(* IEC 61131-3 sources: daoli-st-library/DL_Process (part 8) *)

(* ---- FB_DL_TruckScaleSeq.st ---- *)
(*==============================================================================
 * 组件名称 (Component)  : FB_DL_TruckScaleSeq
 * 所属子库 (Sublibrary) : DL_Process
 * 当前版本 (Version)    : 1.0.2
 * 兼容性   (Platform)   : CODESYS 3.5 / TwinCAT 3 / 汇川 InoProShop / Machine Expert
 *                         仅依赖 Standard.library + DL_ 库内既有件，零厂商方言
 * 来源标签 (Source)     : self-std
 * 功能描述 (Function)   : 车辆过磅称重流程七态顺控：空载等待 -> 车辆上磅（到位
 *                         开关）-> 稳定窗（称重稳定判据，委托 FB_DL_SignalStatistics
 *                         统计内核，峰峰值 < 容差判稳）-> 读数锁存（皮重 / 毛重
 *                         配对）-> 下磅 -> 台账推进（8 条定长环形，写指针饱和）。
 *                         超时未稳定置码重测；防作弊窗（读数期间磅台扰动检测）；
 *                         毛重 < 皮重（亏吨）显式码不静默取负净重。
 * 委托清单 (Delegation) : FB_DL_SignalStatistics（DL_MathData，稳态窗口径次源，
 *                         实例化组合调用——峰峰值 fRange 即稳定判据核）
 * 配比约束 (R100)       : tStableTimeout 必须大于统计窗填满耗时（nStableSamples ×
 *                         任务周期），否则未满窗即被超时重测，稳定判据永不达成。
 * 遗留假设三句声明 (R95): ①代理值：稳定窗以「样本数 nStableSamples × 任务周期」
 *                         代理时间窗 tStableWin；②覆盖范围：任务周期已知且恒定的
 *                         调用场合；③覆盖不到的区间：任务周期漂移 / 变长场合由
 *                         tStableTimeout 超时重测兜底，最坏表现是判稳变慢而非误判。
 * 边界与语义披露 (Boundary disclosure) :
 *   1) 读数未锁存前下磅（bOnScale 在稳定 / 锁存相消失）-> 流程作废 + 台账不写入
 *      （信息级），统计窗清零重来。
 *   2) 防作弊窗：稳定相内磅台到位信号闪断视为扰动（车未完全上磅 / 人为干预），
 *      置信息级并回稳定相重测，杜绝在扰动读数上锁存。
 *   3) 毛重 < 皮重（亏吨）为显式信息级：净重置 0 出台账，绝不静默取负
 *      （负净重会污染库存对账，R81 还原方向不饱和口径同理）。
 *   4) 皮 / 毛配对以「皮重槽与毛重槽均已锁存」为准，不做车号强校验（车号仅入
 *      台账留痕）；配对完成后双槽清零迎接下一车。
 *   5) 称重值非有限属**运行时信号失效**，不是组态错误：自 v1.0.2 起拆为独立信号闸——
 *      本拍只判 NaN / Inf 并置信息级 16#0005_04DD，统计与判据一律使用上一次有效值
 *      快照（fWeightHold），不锁存、不置 bError、不迁 eFault；失效持续由稳定超时
 *      重测（04D9）兜底。判定拍与消费拍强制错开一拍（本拍判定 -> 下拍消费
 *      bWeightBad），杜绝同拍把脏值锁进皮毛槽。
 *   6) 组态闸（bCfgBad）自 v1.0.2 起只含**静态组态量**（容差 / 超时窗 / 窗样本数），
 *      运行时信号不得进入组态锁存路径（避免一拍 NaN 让磅房永久锁死，R152）。
 * 故障码表 (Error codes) :
 *   16#0005_03B2 [故障级] 稳定窗组态非法（容差 <= 0 / 超时 <= 0 / 窗样本数越域）
 *                 反证：回退后流程照常，码位是组态错误唯一可见出口。
 *   16#0005_04D6 [信息级] 未锁存先下磅，流程作废台账不写入
 *                 反证：作废后回空闲与「正常完成」输出组合不同但作废原因（司机
 *                 误操作 / 磅台故障）不可区分，码位承载事件事实。
 *   16#0005_04D7 [信息级] 亏吨（毛重 < 皮重），净重置 0 出台账
 *                 反证：净重 0 与「空车皮重恰好等于毛重」组合相同，码位区分
 *                 正常零载与亏吨异常。
 *   16#0005_04D8 [信息级] 读数期磅台扰动（防作弊窗触发），重测
 *                 反证：重测与「正常重来」输出组合相同，码位是防作弊事实唯一出口。
 *   16#0005_04D9 [信息级] 超时未稳定，清窗重测
 *                 反证：重测与防作弊重测输出组合相似（均回稳定相），码位区分
 *                 「称量不稳」与「磅台扰动」两种成因（R190）。
 *   16#0005_04DD [信息级] 称重信号非有限（NaN / Inf），保持上次有效值不锁存
 *                 反证：保持时 fWeightHold 不变，与「称重值恰好稳定不变」的输出组合
 *                 完全相同；无码则信号断线被误读为「读数极稳」而照常判稳锁存，
 *                 该误判在现有输出上不可观测（R90 反证成立，R69 点修④）。
 * 码位总账 (Code ledger) : 16#0005_03B2 用 ｜ 16#0005_04D6 / 04D7 / 04D8 / 04D9 / 04DD 用
 * 依赖     (Depends)    : FB_DL_SignalStatistics
 * 红线自检 (Redline)    : R1 ✓ 零全局变量与 VAR_EXTERNAL ｜ R2 ✓ 零 %I/%Q 物理地址
 *                         R3 ✓ 纯 IEC 61131-3 + 库内委托件
 *                         R4 ✓ 域闸全枚举 / 计数饱和 / 浮点容差比较（fRange < 容差直比）
 *                         R5 ✓ 全变量中英双语同行注释 ｜ R6 ✓ 七态 ENUM + CASE + ELSE 兜底
 *                         R7 ✓ 二沿二计时 + 统计委托件每拍无条件调用
 * 修订历史 (Revision)   :
 *   2026-11-22  v1.0.0  首版入库（R68 构建轮 · 批 3 · 目标 15）
 *   2026-11-22  v1.0.1  终审就地修①②③：组态锁存解除路径可达化 + 超时重测清窗单拍化 + 皮毛槽镜像输出复核
 *   2026-11-22  v1.0.2  R69 点修④：称重信号非有限（NaN）自组态闸拆出为独立信号闸——判定与
 *                       消费分两拍（本拍判 NaN 只置标志与信息码，下一拍才作用于判稳与挂起），
 *                       失效期保持上次有效值、不锁存、不置 bError
 *============================================================================*)

(*-----------------------------------------------------------------------------
 * 枚举: E_DL_ScaleSeqState（归属 DL_Process，与 FB_DL_TruckScaleSeq 同文件）
 *----------------------------------------------------------------------------*)
TYPE E_DL_ScaleSeqState :
(
    eIdle      := 0,    // 空载等待：无车在磅 / Idle, no truck on scale
    eOnScale   := 10,   // 车辆上磅确认：到位保持 / Truck on scale, arrival confirmed
    eStabilize := 20,   // 稳定窗：统计判稳 / Stabilising, statistics window
    eLatch     := 30,   // 读数锁存：皮 / 毛配对 / Latching, tare-gross pairing
    eOffScale  := 40,   // 下磅：等车辆离开 / Off scale, waiting for departure
    eDone      := 50,   // 台账推进完成拍 / Ledger advanced, one-shot
    eFault     := 99    // 组态锁存：流程拒绝 / Config latched, flow refused
);
END_TYPE

(*==============================================================================
 * 功能块: FB_DL_TruckScaleSeq
 * 调用约定: 每个扫描周期无条件调用一次；bOnScale / bTareMode 为电平引脚。
 *============================================================================*)
FUNCTION_BLOCK FB_DL_TruckScaleSeq
VAR_INPUT
    fWeight       : REAL;                // 磅台称重值 [kg] / Scale weight [kg]
    bOnScale      : BOOL;                // 磅台到位开关（车辆在磅）/ Truck-on-scale limit switch
    bTareMode     : BOOL;                // 本次称量模式：TRUE = 皮重 / TRUE tare, FALSE gross
    uTruckId      : UINT;                // 车号 [号]，仅入台账留痕 / Truck id, ledger only
    nStableSamples: INT  := 32;          // 稳定统计窗样本数 [个]，域 2..64 / Stability window samples
    fStableTolKg  : REAL := 50.0;        // 稳定判据峰峰值容差 [kg] / Stability peak-to-peak tolerance [kg]
    tStableTimeout: TIME := T#30S;       // 稳定超时窗 [s]，须宽于窗填满耗时 / Stability timeout [s]
    bEnable       : BOOL := TRUE;        // 使能 / Enable
    bReset        : BOOL;                // 上升沿：清组态锁存与台账计数 / Rising edge: clear latches
END_VAR
VAR_OUTPUT
    eState       : E_DL_ScaleSeqState;   // 当前状态（供 HMI 诊断）/ Current state
    fTareLatched : REAL;                 // 当前皮重槽 [kg]，0 = 未锁存 / Current tare slot, 0 = unset
    fGrossLatched: REAL;                 // 当前毛重槽 [kg]，0 = 未锁存 / Current gross slot, 0 = unset
    fNetLast     : REAL;                 // 最近一票净重 [kg] / Last net weight [kg]
    nLedgerCount : INT;                  // 台账有效票数 [票]，0..8 / Ledger entry count
    bLedgerFull  : BOOL;                 // 台账已满回卷（最旧被覆盖）/ Ledger full, oldest overwritten
    bJudgeSuspended : BOOL;              // 稳定判据挂起（窗未满 / 称重值无效）/ Judge suspended
    bError       : BOOL;                 // 故障标志（组态锁存）/ Fault flag
    uErrorId     : UDINT;                // 故障码，0 = 无故障 / Error code, 0 = none
END_VAR
VAR
    fbTrigReset  : R_TRIG;               // 复位沿检测实例 / Reset edge detector
    fbTrigOn     : R_TRIG;               // 上磅沿检测实例 / On-scale edge detector
    tonStableTo  : TON;                  // 稳定超时计时实例 / Stability timeout timer
    fbStat       : FB_DL_SignalStatistics; // 统计委托实例 / Statistics delegate
    eStateInt    : E_DL_ScaleSeqState;   // 主状态机内部当前态 / Internal state machine state
    auiTruck     : ARRAY[0..7] OF UINT;  // 台账车号环形 [号] / Ledger truck id ring
    afTareRing   : ARRAY[0..7] OF REAL;  // 台账皮重环形 [kg] / Ledger tare ring [kg]
    afGrossRing  : ARRAY[0..7] OF REAL;  // 台账毛重环形 [kg] / Ledger gross ring [kg]
    afNetRing    : ARRAY[0..7] OF REAL;  // 台账净重环形 [kg] / Ledger net ring [kg]
    nLedgerWrite : INT;                  // 台账写指针 [0..7] / Ledger write pointer
    uLedgerTotal : UDINT;                // 台账累计票数 [票]（回卷判据）/ Ledger total ever
    fTareInt     : REAL;                 // 皮重槽内部副本 [kg] / Internal tare slot
    fGrossInt    : REAL;                 // 毛重槽内部副本 [kg] / Internal gross slot
    fWeightSnap  : REAL;                 // 锁存读数快照 [kg] / Latched weight snapshot
    fWeightHold  : REAL;                 // 上次有效称重值快照 [kg]（信号失效期供统计）/ Last valid weight snapshot [kg]
    bWeightBadT  : BOOL;                 // 本拍称重信号非有限（NaN / Inf）/ Weight non-finite this scan
    bWeightBad   : BOOL;                 // 滞后一拍的信号失效标志（消费用）/ Delayed signal-invalid flag for consumption
    nWinEff      : INT;                  // 钳位后窗样本数 [个] / Clamped window samples
    fTolEff      : REAL;                 // 钳位后容差 [kg] / Clamped tolerance
    bStatClear   : BOOL;                 // 统计窗清零脉冲（单拍）/ Statistics clear pulse
    bCfgBad      : BOOL;                 // 本拍组态非法 / Config illegal this scan
    bCfgLatch    : BOOL;                 // 组态故障锁存 / Config fault latch
    bErrorInt    : BOOL;                 // 本拍故障置位累加（出口归并）/ Fault set accumulator
    bToutPulse   : BOOL;                 // 超时清窗单拍已发标志（防每拍清窗死循环）/ Timeout clear issued flag
    bFirstScan   : BOOL := TRUE;         // 上电首扫标志 / First-scan flag
END_VAR
VAR CONSTANT
    DL_TS_WIN_MIN  : INT  := 2;      // 窗样本数下限 [个]（统计件域）/ Window floor
    DL_TS_WIN_MAX  : INT  := 64;     // 窗样本数上限 [个]（统计件域）/ Window ceiling
    DL_TS_LEDGER   : INT  := 8;      // 台账深度 [票] / Ledger depth
    DL_TS_FIN_LIM  : REAL := 1.0E30; // REAL 有限幅值判界 / REAL finiteness bound
END_VAR

(*------------------------------------------------------------------------------
 * 段 1｜无条件刷新区（红线 R7）：二沿一计时 + 统计委托件每拍调用
 *      Unconditional refresh: two edges, one timer, the stats delegate every scan
 *-----------------------------------------------------------------------------*)
fbTrigReset(CLK := bReset);
fbTrigOn(CLK := bOnScale);
tonStableTo(IN := (eStateInt = E_DL_ScaleSeqState.eStabilize), PT := tStableTimeout);

fbStat(fIn := fWeightHold, bSample := TRUE, nWindow := nWinEff, bClear := bStatClear);

(*------------------------------------------------------------------------------
 * 段 2｜上电首扫：台账与配对槽显式落零
 *      First-scan init: ledger and pairing slots cleared explicitly
 *-----------------------------------------------------------------------------*)
IF bFirstScan THEN
    eStateInt    := E_DL_ScaleSeqState.eIdle;
    fTareInt     := 0.0;
    fGrossInt    := 0.0;
    fWeightSnap  := 0.0;
    fWeightHold  := 0.0;                 // 保持槽首扫落零 [kg] / Hold slot cleared on first scan
    bWeightBad   := FALSE;               // 滞后失效标志首扫落假 / Delayed invalid flag cleared
    nLedgerWrite := 0;
    uLedgerTotal := 0;
    bFirstScan   := FALSE;
END_IF

(*------------------------------------------------------------------------------
 * 段 3｜每拍预清（FB32-1）：单拍标志，禁入锁存 / 快照 / 台账
 *      Per-scan preset: single-scan flags only
 *-----------------------------------------------------------------------------*)
bErrorInt  := FALSE;
bStatClear := FALSE;

(*------------------------------------------------------------------------------
 * 段 4｜组态域闸（R151 全枚举）+ 两级回退（R117）
 *      Config gate with two-level fallback
 *      解除路径（R152 自证）：复位沿 AND 组态改对
 *      R69 点修④：组态闸只含静态组态量；称重信号非有限一律不进本闸（见段 4b）
 *-----------------------------------------------------------------------------*)
bCfgBad := (fStableTolKg <= 0.0) OR (fStableTolKg <> fStableTolKg)
           OR (tStableTimeout <= T#0S)
           OR (nStableSamples < DL_TS_WIN_MIN) OR (nStableSamples > DL_TS_WIN_MAX);

IF bCfgBad THEN
    bCfgLatch := TRUE;
END_IF

IF (fStableTolKg <= 0.0) OR (fStableTolKg <> fStableTolKg) THEN
    fTolEff := 50.0;                 // 回退默认容差 / Fallback default tolerance
ELSE
    fTolEff := fStableTolKg;         // 合法直通 / Valid pass-through
END_IF

IF (nStableSamples < DL_TS_WIN_MIN) OR (nStableSamples > DL_TS_WIN_MAX) THEN
    nWinEff := 32;                   // 回退默认窗长 / Fallback default window
ELSE
    nWinEff := nStableSamples;       // 合法直通 / Valid pass-through
END_IF

IF bCfgLatch THEN
    uErrorId  := 16#0005_03B2;       // 故障级：稳定窗组态非法 / Fault: config illegal
    bErrorInt := TRUE;
END_IF

(* 终审就地修 v1.0.1（R68①②）：解除路径（R152 自证可达）——复位沿 AND 组态非法
 * 条件消失即清锁存。原实现把组态锁存清零只写在 eFault 相分支，而组态闸置锁存后
 * 不迁相（只回 eIdle 驻留），eFault 相不可达 -> 锁存永不可解，磅房流程一次性
 * 永久死锁至 PLC 重启（终审两式①）。 *)
IF fbTrigReset.Q AND (NOT bCfgBad) THEN
    bCfgLatch := FALSE;              // 锁存解除 / Latch cleared
    uErrorId  := 16#0000_0000;       // 码位随解除归零 / Code cleared with the latch
END_IF

(*------------------------------------------------------------------------------
 * 段 4b｜信号闸（R69 点修④）：非有限只判不锁，判定拍与消费拍强制错开一拍
 *      Signal gate: non-finite is judged here and consumed one scan later
 *      拍 N：本拍判 bWeightBadT（NaN 自反 + Inf 差自减 + 幅值兜底），失效即置信息码
 *            04DD，**不写** fWeightHold、不锁存、不迁相；
 *      拍 N+1：bWeightBad 才被统计判据与 bJudgeSuspended 消费（错开一拍，防同拍
 *            把脏值锁进皮毛槽 / 判稳窗）。
 *-----------------------------------------------------------------------------*)
bWeightBadT := (fWeight <> fWeight)
               OR ((fWeight - fWeight) <> (fWeight - fWeight))
               OR (ABS(fWeight) >= DL_TS_FIN_LIM);
IF bWeightBadT THEN
    uErrorId := 16#0005_04DD;        // 信息级：信号非有限，保持上次有效值 / Info: non-finite, holding last valid
ELSE
    fWeightHold := fWeight;          // 有效样本刷新保持槽 [kg] / Refresh the hold slot with a valid sample
END_IF
(* 消费侧滞后镜像 bWeightBad 在主体末行统一刷新（见段 7 之后），保证「本拍判定、
 * 下拍消费」两拍分离，CASE 与判稳判据读到的永远是上一拍结论。 *)
(* The mirror bWeightBad is refreshed on the last body line, so every consumer reads the previous verdict *)

(*------------------------------------------------------------------------------
 * 段 5｜主状态机（红线 R6）：ENUM + CASE + ELSE 兜底
 *      Main state machine with the mandatory ELSE fallback
 *      同拍竞态（R275）：锁存相先消化本拍锁存，再消化下磅沿
 *-----------------------------------------------------------------------------*)
CASE eStateInt OF

    E_DL_ScaleSeqState.eIdle:
        IF bCfgLatch OR (NOT bEnable) THEN
            (* 组态 / 失能驻留：流程拒绝（降级语义已声明）/ Flow refused, declared *)
        ELSIF fbTrigOn.Q THEN
            bStatClear := TRUE;      // 新车进窗先清统计 / Clear stats for the new truck
            eStateInt  := E_DL_ScaleSeqState.eOnScale;
        END_IF

    E_DL_ScaleSeqState.eOnScale:
        IF NOT bOnScale THEN
            (* 读数未锁存前下磅：流程作废 + 台账不写入（信息级 0405） *)
            (* Departure before any latch: flow voided, ledger untouched *)
            bStatClear := TRUE;
            uErrorId   := 16#0005_04D6;   // 信息级：未锁存先下磅 / Info: departed unlatched
            eStateInt  := E_DL_ScaleSeqState.eIdle;
        ELSE
            eStateInt := E_DL_ScaleSeqState.eStabilize;   // 到位保持确认，进稳定窗 / Confirmed, to stabilise
        END_IF

    E_DL_ScaleSeqState.eStabilize:
        IF (NOT bOnScale) AND (NOT fbTrigOn.Q) THEN
            (* 防作弊窗：稳定相内到位信号消失 = 扰动（车未完全上磅 / 人为干预） *)
            (* Anti-cheat: on-scale dropped during stabilising is a disturbance *)
            bStatClear := TRUE;      // 清窗重测 / Clear and re-measure
            uErrorId   := 16#0005_04D8;   // 信息级：磅台扰动 / Info: disturbance
            eStateInt  := E_DL_ScaleSeqState.eIdle;   // 作废回空闲（未锁存不写台账）/ Voided
        ELSIF (fbStat.nCount >= nWinEff) AND (fbStat.fRange < fTolEff) THEN
            eStateInt := E_DL_ScaleSeqState.eLatch;   // 窗满且峰峰值达标 / Full window, range OK
        END_IF

    E_DL_ScaleSeqState.eLatch:
        IF (fWeight <> fWeight) OR ((fWeight - fWeight) <> (fWeight - fWeight))
           OR (ABS(fWeight) >= DL_TS_FIN_LIM) OR bWeightBad THEN
            (* 称重值非有限：拒绝锁存（保持槽不写），回稳定相由超时兜底 *)
            (* Non-finite weight: latch refused, back to stabilise *)
            bStatClear := TRUE;
            eStateInt  := E_DL_ScaleSeqState.eStabilize;
        ELSE
            fWeightSnap := fWeight;  // 读数锁存 / Latch the reading
            IF bTareMode THEN
                fTareInt := fWeightSnap;      // 皮重入槽 / Tare into slot
            ELSE
                fGrossInt := fWeightSnap;     // 毛重入槽 / Gross into slot
            END_IF
            IF (fTareInt > 0.0) AND (fGrossInt > 0.0) THEN
                WriteLedger();       // 皮毛双槽齐 -> 台账（私有方法）/ Pair complete, ledger write
            END_IF
            eStateInt := E_DL_ScaleSeqState.eOffScale;
        END_IF

    E_DL_ScaleSeqState.eOffScale:
        IF NOT bOnScale THEN
            eStateInt := E_DL_ScaleSeqState.eDone;   // 车辆离开 / Truck departed
        END_IF

    E_DL_ScaleSeqState.eDone:
        eStateInt := E_DL_ScaleSeqState.eIdle;       // 单拍完成相：下一拍回空闲 / One-shot, back to idle

    E_DL_ScaleSeqState.eFault:
        IF fbTrigReset.Q AND (NOT bCfgBad) THEN
            bCfgLatch := FALSE;      // 解除路径自证可达（R152）/ Clear path reachable
            uErrorId  := 16#0000_0000;
            eStateInt := E_DL_ScaleSeqState.eIdle;
        END_IF

    ELSE
        eStateInt := E_DL_ScaleSeqState.eFault;
        uErrorId  := 16#0005_03B2;
        bErrorInt := TRUE;

END_CASE;

(*------------------------------------------------------------------------------
 * 段 6｜超时未稳定消化：清窗重测（信息级），与防作弊重测成因码位互异（R190）
 *      Stability timeout: clear and re-measure, cause code distinct from 0407
 *-----------------------------------------------------------------------------*)
(* 终审就地修 v1.0.1（R68③）：超时重测单拍化。TON.Q 在 IN 保持期间恒真，原实现
 * 每拍 bStatClear := TRUE，统计窗被扫描周期级反复清零 -> 窗永不填满、判稳永不
 * 达成（超时同源挂死）。改为「一次超时只清一次窗」，重测窗得以重新累计。
 * Timeout clear is now a one-shot: an expired timer no longer wipes the window every scan. *)
IF tonStableTo.Q AND (eStateInt = E_DL_ScaleSeqState.eStabilize) AND (NOT bToutPulse) THEN
    bStatClear := TRUE;              // 清窗重测（单拍）/ Clear and re-measure, once
    uErrorId   := 16#0005_04D9;      // 信息级：超时重测 / Info: timeout re-measure
    bToutPulse := TRUE;              // 单拍标志置位 / Mark the one-shot as issued
END_IF
IF eStateInt <> E_DL_ScaleSeqState.eStabilize THEN
    bToutPulse := FALSE;             // 离开稳定相即撤销（下次进相可再清一次）/ Re-armed on phase exit
END_IF

(*------------------------------------------------------------------------------
 * 段 7｜输出单一出口（范式 P-05）：台账口径与挂起标志派生
 *      Single output exit: ledger derived values and the suspension flag
 *-----------------------------------------------------------------------------*)
IF uLedgerTotal > UDINT#8 THEN
    bLedgerFull := TRUE;             // 回卷覆盖（最旧被覆盖）/ Ring wrapped
END_IF
IF UDINT_TO_DINT(uLedgerTotal) < DINT#8 THEN
    nLedgerCount := DINT_TO_INT(UDINT_TO_DINT(uLedgerTotal));
ELSE
    nLedgerCount := 8;               // 深度即上限 [票] / Depth is the cap
END_IF

fTareLatched  := fTareInt;           // 皮重槽镜像输出（0 = 未锁存）/ Mirror tare slot out
fGrossLatched := fGrossInt;          // 毛重槽镜像输出（0 = 未锁存）/ Mirror gross slot out

bJudgeSuspended := (fbStat.nCount < nWinEff) OR bWeightBad
                   OR (eStateInt <> E_DL_ScaleSeqState.eStabilize);

bError := bErrorInt OR (eStateInt = E_DL_ScaleSeqState.eFault);
eState := eStateInt;
bWeightBad := bWeightBadT;           // 主体末行刷新滞后镜像（判定 -> 消费相隔一拍）/ Last line, one-scan delayed mirror
END_FUNCTION_BLOCK

(*------------------------------------------------------------------------------
 * 私有方法: WriteLedger —— 皮 / 毛配对台账唯一写入点（环形 + 写指针饱和）
 *      Private method: the single ledger write, ring with saturating pointer
 *      调用约定: 仅在 eLatch 相皮毛双槽齐拍调用一次；亏吨显式码在此落账
 *----------------------------------------------------------------------------*)
METHOD WriteLedger
VAR
    fNet : REAL;                     // 本票净重 [kg] / Net weight of this ticket
END_VAR

IF fGrossInt >= fTareInt THEN
    fNet := fGrossInt - fTareInt;    // 正常净重 / Normal net
ELSE
    fNet := 0.0;                     // 亏吨：净重置 0 不出负值（R81 口径）/ Tare exceeds gross: zero
    uErrorId := 16#0005_04D7;        // 信息级：亏吨 / Info: negative net
END_IF

auiTruck[nLedgerWrite]   := uTruckId;      // 车号入账 / Truck id into ledger
afTareRing[nLedgerWrite] := fTareInt;      // 皮重入账 / Tare into ledger
afGrossRing[nLedgerWrite] := fGrossInt;    // 毛重入账 / Gross into ledger
afNetRing[nLedgerWrite]  := fNet;          // 净重入账 / Net into ledger

fNetLast    := fNet;               // 最近净重出口留影 / Snapshot last net
fTareInt    := 0.0;                // 配对槽清零迎下一车 / Pair slots cleared
fGrossInt   := 0.0;

uLedgerTotal := uLedgerTotal + 1;  // 累计票数推进（回卷判据）/ Total tickets up
nLedgerWrite := nLedgerWrite + 1;  // 写指针推进 / Pointer up
IF nLedgerWrite >= DL_TS_LEDGER THEN
    nLedgerWrite := 0;              // 显式回卷 / Explicit wrap
END_IF

END_METHOD

(* ---- FC_DL_CathodeCapacityFadeCalc.st ---- *)
(*
  Component : FC_DL_CathodeCapacityFadeCalc
  Category  : DL_Process
  Function  : 容量衰减 = 1 − Qn/Q0，并按模型选择给出线性或平方根预测衰减
  Complexity: C2
  开源溯源 : DLF 内部原创（R94 族模板派生）；参考语义来源见 SOURCE_HUNTING_MATRIX.md
  规则遵从 : R1-R16
  契约     : 输入 rQ0Ah 初始容量 [Ah]、rQnAh 第 n 圈容量 [Ah]、nCycles 循环圈数 [圈]、
             rFadePerCyclePct 线性模型每圈衰减率 [%/圈]、rSqrtCoefPct 平方根模型系数 [%/圈^0.5]、
             eModel 模型选择枚举；输出 rFadePct 实测衰减 [%]、rFadePredPct 模型预测衰减 [%]、
             xValid 有效标志、nFaultCode 故障码。
  边界     : 初始容量为分母须 >1.0E-9 [Ah]；圈数须 ≥1；两个模型系数须 ≥0；
             平方根模型用 SQRT(圈数) 实现，禁用幂运算方言；模型枚举未知值走 ELSE 兜底判 9803。
  码位     : 9801 输入非有限（故障级）；9802 初始容量或圈数非法（故障级）；9803 模型枚举未知或系数越域（故障级）。
*)
TYPE E_DL_CathodeFadeModel :
(
    eLinear := 0,    // 线性衰减模型：fade = k × n EN: the linear fade model
    eSqrt   := 1     // 平方根衰减模型：fade = c × √n EN: the square root fade model
);
END_TYPE

FUNCTION FC_DL_CathodeCapacityFadeCalc : BOOL
VAR_INPUT
    rQ0Ah          : LREAL := 5.0;     // 初始容量 [Ah] EN: the initial capacity of the cell
    rQnAh          : LREAL := 4.5;     // 第 n 圈容量 [Ah] EN: the capacity after the given number of cycles
    nCycles        : INT := 500;       // 循环圈数 [圈] EN: the number of cycles applied
    rFadePerCyclePct: LREAL := 0.02;   // 线性模型每圈衰减率 [%/圈] EN: the per cycle fade rate of the linear model
    rSqrtCoefPct   : LREAL := 0.4;     // 平方根模型系数 [%/圈^0.5] EN: the coefficient of the square root model
    eModel         : E_DL_CathodeFadeModel;   // 衰减模型选择 [-] EN: the fade model selection
END_VAR
VAR_OUTPUT
    rFadePct     : LREAL;              // 实测容量衰减 [%] EN: the measured capacity fade
    rFadePredPct : LREAL;              // 模型预测容量衰减 [%] EN: the capacity fade predicted by the selected model
    xValid       : BOOL;               // 输出可信标志 EN: the outputs are valid
    nFaultCode   : INT;                // 0=无故障 9801=输入非有限 9802=初始容量或圈数非法 9803=模型或系数越域 EN: zero none, 9801 non finite, 9802 capacity or cycles illegal, 9803 model or coefficient out of range
END_VAR
VAR
    xFinAll : BOOL;                    // 浮点入参同时有限 EN: the floating inputs are finite
    rDen    : LREAL;                   // 分母（初始容量） [Ah] EN: the divisor, the initial capacity
    rFade   : LREAL;                   // 实测衰减中间值 [%] EN: the interim measured fade
    rPred   : LREAL;                   // 预测衰减中间值 [%] EN: the interim predicted fade
    rN      : LREAL;                   // 圈数的实数形式 [圈] EN: the cycle count as a real number
    rSqrtN  : LREAL;                   // 圈数平方根 [圈^0.5] EN: the square root of the cycle count
END_VAR
VAR CONSTANT
    DL_CCF_Z        : LREAL := 0.0;    // 浮点零常量 EN: the floating point zero constant
    DL_CCF_ONE      : LREAL := 1.0;    // 浮点壹常量 EN: the floating point one constant
    DL_CCF_HUNDRED  : LREAL := 100.0;  // 百分数换算系数 EN: the percent conversion factor
    DL_CCF_MIN      : LREAL := 1.0E-9; // 分母绝对值下限 [Ah] EN: the lower bound of the divisor magnitude
    DL_CCF_C_BAD    : INT := 9801;     // 输入非有限 EN: a non finite input
    DL_CCF_C_DEN    : INT := 9802;     // 初始容量或圈数非法 EN: the initial capacity or the cycle count is illegal
    DL_CCF_C_MODEL  : INT := 9803;     // 模型或系数越域 EN: the model or the coefficient is out of range
END_VAR

// 段1｜出口预置
FC_DL_CathodeCapacityFadeCalc := FALSE;   // 返回值预置假 EN: preset the return value to false
rFadePct := DL_CCF_Z;                     // 实测衰减预置零 [%] EN: preset the measured fade to zero
rFadePredPct := DL_CCF_Z;                 // 预测衰减预置零 [%] EN: preset the predicted fade to zero
xValid := FALSE;                          // 有效标志预置假 EN: preset the validity flag to false
nFaultCode := 0;                          // 故障码预置零 EN: preset the fault code to zero

// 段2｜非有限闸：浮点入参全列（两模型系数参与换算，漏则模型输出可为 NaN）
xFinAll := (rQ0Ah = rQ0Ah) AND ((rQ0Ah - rQ0Ah) = DL_CCF_Z)
        AND (rQnAh = rQnAh) AND ((rQnAh - rQnAh) = DL_CCF_Z)
        AND (rFadePerCyclePct = rFadePerCyclePct) AND ((rFadePerCyclePct - rFadePerCyclePct) = DL_CCF_Z)
        AND (rSqrtCoefPct = rSqrtCoefPct) AND ((rSqrtCoefPct - rSqrtCoefPct) = DL_CCF_Z);   // 四浮点输入有限性 EN: the finiteness of the four floating inputs
IF NOT xFinAll THEN                                                                          // 非有限出口 EN: leave early on a non finite input
    nFaultCode := DL_CCF_C_BAD;                                                              // 非有限码 EN: the non finite code
    RETURN;                                                                                  // 早退 EN: return early
END_IF

// 段3｜域闸：初始容量过分母下限、圈数 ≥1、容量非负、系数非负
rDen := rQ0Ah;                                                                               // 取分母 [Ah] EN: take the divisor
IF (ABS(rDen) < DL_CCF_MIN) OR (nCycles < 1) OR (rQnAh < DL_CCF_Z) THEN                      // 容量与圈数闸 EN: the capacity and cycle gate
    nFaultCode := DL_CCF_C_DEN;                                                              // 非法码 EN: the illegal code
    RETURN;                                                                                  // 早退 EN: return early
END_IF
IF (rFadePerCyclePct < DL_CCF_Z) OR (rSqrtCoefPct < DL_CCF_Z) THEN                           // 模型系数闸 EN: the model coefficient gate
    nFaultCode := DL_CCF_C_MODEL;                                                            // 系数越域码 EN: the coefficient code
    RETURN;                                                                                  // 早退 EN: return early
END_IF

// 段4｜实测衰减：fade = (1 − Qn/Q0) × 100，不钳位（负衰减表达容量回升，方向信息保留）
rFade := (DL_CCF_ONE - (rQnAh / rDen)) * DL_CCF_HUNDRED;                                     // 实测衰减 [%] EN: the measured fade

// 段5｜模型预测：ENUM + CASE 且 ELSE 兜底
rN := INT_TO_LREAL(nCycles);                                                                 // 圈数转实数 [圈] EN: the cycle count as a real number
CASE eModel OF
    E_DL_CathodeFadeModel.eLinear:
        rPred := rFadePerCyclePct * rN;                                                      // 线性模型 [%] EN: the linear model
    E_DL_CathodeFadeModel.eSqrt:
        rSqrtN := SQRT(rN);                                                                  // 圈数平方根，圈数已证 ≥1 [圈^0.5] EN: the square root, the count is proven at least one
        rPred := rSqrtCoefPct * rSqrtN;                                                      // 平方根模型 [%] EN: the square root model
ELSE
    nFaultCode := DL_CCF_C_MODEL;                                                            // 未知模型码 EN: the unknown model code
    rFadePct := rFade;                                                                       // 实测值仍可给出 [%] EN: the measured value is still published
    RETURN;                                                                                  // 早退 EN: return early
END_CASE

// 段6｜结果复检与出口
IF (rFade <> rFade) OR (rPred <> rPred) THEN                                                 // 复检：两路输出非有限 EN: recheck both outputs for a non finite value
    nFaultCode := DL_CCF_C_MODEL;                                                            // 复检失败码 EN: the recheck failure code
    RETURN;                                                                                  // 早退，出口保持零哨兵 EN: return early with the zero sentinels
END_IF
rFadePct := rFade;                                                                           // 实测衰减出口 [%] EN: the measured fade output
rFadePredPct := rPred;                                                                       // 预测衰减出口 [%] EN: the predicted fade output
xValid := TRUE;                                                                              // 结果可信 EN: the results are valid
FC_DL_CathodeCapacityFadeCalc := TRUE;                                                       // 返回真 EN: return true
END_FUNCTION

(* ---- FC_DL_AirCompFreeAirDeliveryCalc.st ---- *)
(*
  Name: FC_DL_AirCompFreeAirDeliveryCalc
  Category: DL_Process
  Version: 1.0.0
  Round: R90 / 2026-11-25
  开源溯源：clean-room 自研（族 压缩空气系统能效，ST 开源生态实测 0 命中，无外部代码引入）
  功能：1) 储气罐压降法测自由排气量 FAD：空压机向储气罐充气（或罐内气体对外供气）期间，
           罐内绝对压降对应的「常压自由空气容积」= 罐容积 × 压降 / 大气压，
           再按测量时长折算到每分钟即得 FAD：fFadM3min = V_tank · ΔP / P_atm · 60 / t。
           该法假设过程等温（罐体与外界充分换热），适用于离线产能测试。
        2) 标准状态折算：把实测工况（fTempC、fAtmBar）下的自由空气折算到 0 °C、1013.25 mbar
           的标准状态，用于跨季节、跨海拔的产能对比：fFadNorm = fFad · (273.15/(273.15+t)) · (P_atm/P_std)。
           温度项与压力项均为无因次比值，且方向相反（温度升高使标准容积变小、压力升高使其变大）。
  边界条件：1) 非有限值闸：五路实值入参统一过 NOT(x > -DL_BIG AND x < DL_BIG)，
           同时拦 NaN 与 Inf，命中即拦断实值通路（两个 REAL 输出强制 0.0）并置无效（R19）。
        2) 分母零闸：ABS(fTimeS) > DL_EPS（测量时长为 0 则流速发散）与
           ABS(fAtmBar) > DL_EPS（大气压为 0 则折算无意义）都必须通过，否则判无效。
        3) 开尔文偏移零闸：fTempC 必须 > DL_K0_NEG（−273.15 °C）之上，否则 273.15 + t 为 0 或负，
           标准状态折算的温度分母发散；同时对温度做 −50 ~ 80 °C 的工况量程校验，越域判无效。
        4) 负值与零压降：罐容积为负、压降为负（压力反向上升）均判无效；
           压降为 0 属合法但无信息（FAD = 0），不判无效，仅输出 0。
        5) 饱和钳制：FAD 与标准 FAD 结果均钳到 0 ~ DL_FAD_MAX(10000 m3/min)，
           防测量时长极短导致折算值溢出。
  量纲自证：V·ΔP/P_atm = m3 × bar / bar = m3（自由空气容积，bar 消去）；
           再乘 60 s/min 除 t[s] → m3/min，量纲闭合；
           标准折算两个因子 (K/K) 与 (mbar/mbar) 均为无因次，不改变量纲。
*)

FUNCTION FC_DL_AirCompFreeAirDeliveryCalc : BOOL
VAR_INPUT
    fTankM3       : REAL;   // 储气罐有效容积 [m3] / Effective receiver volume [m3]
    fDropBar      : REAL;   // 测量期间罐内压降 [bar] / Pressure drop during test [bar]
    fTimeS        : REAL;   // 测量时长 [s] / Measurement duration [s]
    fAtmBar       : REAL;   // 当地大气压 [bar] / Local atmospheric pressure [bar]
    fTempC        : REAL;   // 环境温度 [°C] / Ambient temperature [°C]
END_VAR
VAR_OUTPUT
    fFadM3min     : REAL;   // 工况自由排气量 [m3/min] / Free air delivery at site conditions [m3/min]
    fFadNormM3min : REAL;   // 标准状态自由排气量 [m3/min] / Free air delivery at standard conditions
    xValid        : BOOL;   // 计算有效标志 [bool] / Calculation valid flag [bool]
END_VAR
VAR
    _fFreeVolumeM3: REAL;   // 压降对应的常压自由空气容积 [m3] / Free air volume from pressure drop [m3]
    _fFadRawM3min : REAL;   // 未饱和的工况 FAD [m3/min] / Raw site FAD [m3/min]
    _fTempFactor  : REAL;   // 标准状态温度折算因子 [-] / Standard-state temperature factor [-]
    _fPressFactor : REAL;   // 标准状态压力折算因子 [-] / Standard-state pressure factor [-]
    _fNormRawM3min: REAL;   // 未饱和的标准状态 FAD [m3/min] / Raw standard FAD [m3/min]
END_VAR
VAR CONSTANT
    DL_EPS        : REAL := 1.0E-9;    // 分母零闸阈值 [-] / Division-zero gate threshold [-]
    DL_BIG        : REAL := 1.0E12;    // 非有限值闸量级上限 [-] / Finiteness gate magnitude [-]
    DL_K0         : REAL := 273.15;    // 摄氏转开尔文偏移 [K] / Celsius to Kelvin offset [K]
    DL_S_PER_MIN  : REAL := 60.0;      // min → s 换算因子 [s/min] / Minute to second factor [s/min]
    DL_P_STD_MBAR : REAL := 1013.25;   // 标准大气压 [mbar] / Standard atmospheric pressure [mbar]
    DL_T_LO_C     : REAL := -50.0;     // 环境温度量程下限 [°C] / Ambient temperature range low [°C]
    DL_T_HI_C     : REAL := 80.0;      // 环境温度量程上限 [°C] / Ambient temperature range high [°C]
    DL_FAD_MAX    : REAL := 10000.0;   // FAD 饱和钳制上限 [m3/min] / FAD saturation ceiling [m3/min]
END_VAR

(* —— 段 1：非有限值闸（R19：五路入参全覆盖，拦 NaN 与 Inf） —— *)
IF NOT (fTankM3 > -DL_BIG AND fTankM3 < DL_BIG)
   OR NOT (fDropBar > -DL_BIG AND fDropBar < DL_BIG)
   OR NOT (fTimeS > -DL_BIG AND fTimeS < DL_BIG)
   OR NOT (fAtmBar > -DL_BIG AND fAtmBar < DL_BIG)
   OR NOT (fTempC > -DL_BIG AND fTempC < DL_BIG) THEN
    fFadM3min := 0.0;                       // 输出强制 0.0 / Output forced to zero
    fFadNormM3min := 0.0;                   // 标准 FAD 强制 0.0 / Standard FAD forced to zero
    xValid := FALSE;                        // 有效位清零 / Validity cleared
    FC_DL_AirCompFreeAirDeliveryCalc := FALSE;   // 返回码同源 / Return mirrors validity
    RETURN;                                 // 立即退出 / Immediate exit
END_IF

(* —— 段 2：分母零闸（R4：测量时长与大气压两个分母都要闸） —— *)
IF (ABS(fTimeS) <= DL_EPS) OR (ABS(fAtmBar) <= DL_EPS) THEN
    fFadM3min := 0.0;                       // 输出强制 0.0 / Output forced to zero
    fFadNormM3min := 0.0;                   // 标准 FAD 强制 0.0 / Standard FAD forced to zero
    xValid := FALSE;                        // 判无效 / Invalid
    FC_DL_AirCompFreeAirDeliveryCalc := FALSE;   // 返回码同步 / Return synchronised
    RETURN;                                 // 提前退出 / Early exit
END_IF

(* —— 段 3：开尔文偏移零闸与负值闸（温度分母 / 负容积 / 负压降 / 负时长） —— *)
IF ((fTempC + DL_K0) <= DL_EPS)
   OR (fTankM3 < 0.0) OR (fDropBar < 0.0) OR (fTimeS < 0.0) OR (fAtmBar < 0.0) THEN
    fFadM3min := 0.0;                       // 输出强制 0.0 / Output forced to zero
    fFadNormM3min := 0.0;                   // 标准 FAD 强制 0.0 / Standard FAD forced to zero
    xValid := FALSE;                        // 判无效 / Invalid
    FC_DL_AirCompFreeAirDeliveryCalc := FALSE;   // 返回码同步 / Return synchronised
    RETURN;                                 // 提前退出 / Early exit
END_IF

(* —— 段 4：压降法主算式（R22 方向自核：压降越大自由空气越多，除的是大气压不是工况压力） —— *)
_fFreeVolumeM3 := fTankM3 * fDropBar / fAtmBar;                        // 常压自由空气容积 [m3]
_fFadRawM3min := _fFreeVolumeM3 * DL_S_PER_MIN / fTimeS;               // 折算到每分钟 [m3/min]

(* —— 段 5：标准状态折算（温度项与压力项方向相反，均为无因次比值） —— *)
_fTempFactor := DL_K0 / (DL_K0 + fTempC);                              // 温度折算 [-]
_fPressFactor := fAtmBar / (DL_P_STD_MBAR / 1000.0);                   // 压力折算（mbar → bar）[-]
_fNormRawM3min := _fFadRawM3min * _fTempFactor * _fPressFactor;        // 标准状态 FAD [m3/min]

(* —— 段 6：有效位单点聚合（温度工况量程校验） —— *)
xValid := (fTempC >= DL_T_LO_C) AND (fTempC <= DL_T_HI_C)              // 温度在工况量程内
          AND (fTankM3 >= 0.0) AND (fDropBar >= 0.0)                   // 容积与压降非负
          AND (fTimeS > DL_EPS) AND (fAtmBar > DL_EPS);                // 两个分母均为正

(* —— 段 7：输出单点写盘（饱和钳制，防极短测量时长溢出） —— *)
fFadM3min := LIMIT(0.0, _fFadRawM3min, DL_FAD_MAX);                    // 工况 FAD [m3/min]
fFadNormM3min := LIMIT(0.0, _fNormRawM3min, DL_FAD_MAX);               // 标准 FAD [m3/min]
FC_DL_AirCompFreeAirDeliveryCalc := xValid;                            // 返回码：TRUE = 计算可信

END_FUNCTION

(* ---- FC_DL_AirCompLoadUnloadHystCalc.st ---- *)
(*
  Name: FC_DL_AirCompLoadUnloadHystCalc
  Category: DL_Process
  Version: 1.0.0
  Round: R90 / 2026-11-25
  开源溯源：clean-room 自研（族 压缩空气系统能效，ST 开源生态实测 0 命中，无外部代码引入）
  功能：1) 加载/卸载压力带以目标压力为中心对称展开：加载压力 = 目标 − 回差/2，
           卸载压力 = 目标 + 回差/2。两点的间距恰为回差带宽，中心与目标压力重合，
           保证系统的长期平均压力不偏离设定值（若单侧展开会导致平均压力偏移）。
        2) 可行性判定 xViable 由三条独立条件聚合：
             a) 回差带宽不得小于「由最小循环时间反算的最小回差」：把频繁启停的成因归为
                单位时间内压力变化过快，故取经验压力变化速率 DL_RATE_BAR_PER_S 乘最小循环时间
                得到所需回差下限（bar/s × s = bar，量纲闭合），回差低于该下限判不可行；
             b) 储气罐缓冲自由空气容积（罐容积 × 回差 / 大气压）不得低于 DL_BUF_MIN，
                否则回差再大也被小罐吃掉，压力仍会抖动；
             c) 加载压力必须严格为正，否则加载点落到负压区，逻辑上永不加载。
        3) 输出加载/卸载压力供压力开关或控制器组态直接取用。
  边界条件：1) 非有限值闸：四路实值入参统一过 NOT(x > -DL_BIG AND x < DL_BIG)，
           同时拦 NaN 与 Inf，命中即拦断实值通路（两个压力输出强制 0.0、xViable 强制 FALSE）
           并置无效（R19），无效数据不得输出可组态的压力带。
        2) 分母零闸：本件除数仅为常量 2.0 与 DL_P_ATM_BAR，均为常量非零；
           但罐容积必须 > DL_EPS 才能得到有意义的缓冲容积，否则按 0 处理并判不可行。
        3) 负值闸：目标压力为负、回差为负、最小循环时间为负、罐容积为负均判无效
           （回差为负会使加载压力高于卸载压力，压力带反号，属组态错误）。
        4) 零值语义：回差为 0 表示无回差（加载点 = 卸载点，必然频繁启停），
           不判无效但 xViable 必为 FALSE，由可行性判定拦截。
        5) 饱和钳制：目标压力钳 0 ~ DL_P_MAX(40 bar)，回差钳 0 ~ DL_HYST_MAX(10 bar)，
           防组态越界把压力带推到量程外。
  量纲自证：fLoadBar = bar − bar/2 = bar；fUnloadBar = bar + bar/2 = bar，三条均为 bar；
           fHystNeedBar = (bar/s) × (s) = bar，与回差同量纲后方可比较；
           缓冲容积 = m3 × bar / bar = m3。
*)

FUNCTION FC_DL_AirCompLoadUnloadHystCalc : BOOL
VAR_INPUT
    fTargetBar      : REAL;   // 目标压力（压力带中心）[bar] / Target pressure, band centre [bar]
    fHystBar        : REAL;   // 回差带宽 [bar] / Hysteresis band width [bar]
    fMinCycleS      : REAL;   // 允许的最小循环时间 [s] / Minimum allowed cycle time [s]
    fRecvM3         : REAL;   // 储气罐有效容积 [m3] / Effective receiver volume [m3]
END_VAR
VAR_OUTPUT
    fLoadBar        : REAL;   // 加载压力 [bar] / Load pressure [bar]
    fUnloadBar      : REAL;   // 卸载压力 [bar] / Unload pressure [bar]
    fHystNeedBar    : REAL;   // 由最小循环时间反算的最小回差 [bar] / Minimum required hysteresis [bar]
    fBufferM3       : REAL;   // 回差带对应的缓冲自由空气容积 [m3] / Buffer free air volume [m3]
    xViable         : BOOL;   // 压力带可行标志 [bool] / Pressure band feasibility flag [bool]
    xValid          : BOOL;   // 计算有效标志 [bool] / Calculation valid flag [bool]
END_VAR
VAR
    _fTargetClamp   : REAL;   // 钳制后的目标压力 [bar] / Clamped target pressure [bar]
    _fHystClamp     : REAL;   // 钳制后的回差带宽 [bar] / Clamped hysteresis band [bar]
    _fHalfHyst      : REAL;   // 半回差 [bar] / Half hysteresis band [bar]
    _fLoadRawBar    : REAL;   // 未钳制的加载压力 [bar] / Raw load pressure [bar]
    _fUnloadRawBar  : REAL;   // 未钳制的卸载压力 [bar] / Raw unload pressure [bar]
END_VAR
VAR CONSTANT
    DL_EPS          : REAL := 1.0E-9;    // 分母零闸阈值 [-] / Division-zero gate threshold [-]
    DL_BIG          : REAL := 1.0E12;    // 非有限值闸量级上限 [-] / Finiteness gate magnitude [-]
    DL_P_ATM_BAR    : REAL := 1.01325;   // 标准大气压 [bar] / Standard atmospheric pressure [bar]
    DL_P_MAX        : REAL := 40.0;      // 目标压力饱和上限 [bar] / Target pressure saturation ceiling [bar]
    DL_HYST_MAX     : REAL := 10.0;      // 回差带宽饱和上限 [bar] / Hysteresis saturation ceiling [bar]
    DL_RATE_BAR_S   : REAL := 0.0020;    // 经验压力变化速率 [bar/s] / Empirical pressure change rate [bar/s]
    DL_BUF_MIN      : REAL := 0.10;      // 缓冲自由空气容积下限 [m3] / Buffer free air volume lower bound [m3]
    DL_TWO          : REAL := 2.0;       // 半带宽除数（对称展开）[-] / Half-band divisor [-]
END_VAR

(* —— 段 1：非有限值闸（R19：四路入参全覆盖，拦 NaN 与 Inf） —— *)
IF NOT (fTargetBar > -DL_BIG AND fTargetBar < DL_BIG)
   OR NOT (fHystBar > -DL_BIG AND fHystBar < DL_BIG)
   OR NOT (fMinCycleS > -DL_BIG AND fMinCycleS < DL_BIG)
   OR NOT (fRecvM3 > -DL_BIG AND fRecvM3 < DL_BIG) THEN
    fLoadBar := 0.0;                        // 输出强制 0.0 / Output forced to zero
    fUnloadBar := 0.0;                      // 输出强制 0.0 / Output forced to zero
    fHystNeedBar := 0.0;                    // 最小回差强制 0.0 / Minimum hysteresis forced to zero
    fBufferM3 := 0.0;                       // 缓冲容积强制 0.0 / Buffer volume forced to zero
    xViable := FALSE;                       // 可行性强制 FALSE / Feasibility forced off
    xValid := FALSE;                        // 有效位清零 / Validity cleared
    FC_DL_AirCompLoadUnloadHystCalc := FALSE;   // 返回码同源 / Return mirrors validity
    RETURN;                                 // 立即退出 / Immediate exit
END_IF

(* —— 段 2：负值闸（回差为负会使加载压力高于卸载压力，压力带反号） —— *)
IF (fTargetBar < 0.0) OR (fHystBar < 0.0) OR (fMinCycleS < 0.0) OR (fRecvM3 < 0.0) THEN
    fLoadBar := 0.0;                        // 输出强制 0.0 / Output forced to zero
    fUnloadBar := 0.0;                      // 输出强制 0.0 / Output forced to zero
    fHystNeedBar := 0.0;                    // 最小回差强制 0.0 / Minimum hysteresis forced to zero
    fBufferM3 := 0.0;                       // 缓冲容积强制 0.0 / Buffer volume forced to zero
    xViable := FALSE;                       // 可行性强制 FALSE / Feasibility forced off
    xValid := FALSE;                        // 判无效 / Invalid
    FC_DL_AirCompLoadUnloadHystCalc := FALSE;   // 返回码同步 / Return synchronised
    RETURN;                                 // 提前退出 / Early exit
END_IF

(* —— 段 3：饱和钳制（目标压力与回差带宽各自量程） —— *)
_fTargetClamp := LIMIT(0.0, fTargetBar, DL_P_MAX);                // 目标压力钳 0..40 [bar]
_fHystClamp := LIMIT(0.0, fHystBar, DL_HYST_MAX);                 // 回差钳 0..10 [bar]

(* —— 段 4：对称展开压力带（R22 方向自核：加载在下、卸载在上，各偏半个回差） —— *)
_fHalfHyst := _fHystClamp / DL_TWO;                               // 半回差 [bar]
_fLoadRawBar := _fTargetClamp - _fHalfHyst;                       // 加载压力 = 目标 − 半回差 [bar]
_fUnloadRawBar := _fTargetClamp + _fHalfHyst;                     // 卸载压力 = 目标 + 半回差 [bar]

(* —— 段 5：可行性判据量（最小回差 / 缓冲容积） —— *)
fHystNeedBar := DL_RATE_BAR_S * fMinCycleS;                       // bar/s × s = bar
fBufferM3 := fRecvM3 * _fHystClamp / DL_P_ATM_BAR;                // m3 × bar / bar = m3

(* —— 段 6：输出单点写盘（压力带饱和钳制） —— *)
fLoadBar := LIMIT(0.0, _fLoadRawBar, DL_P_MAX);                   // 加载压力钳 0..40 [bar]
fUnloadBar := LIMIT(0.0, _fUnloadRawBar, DL_P_MAX);               // 卸载压力钳 0..40 [bar]

(* —— 段 7：有效位与可行性单点聚合 —— *)
xValid := (fTargetBar >= 0.0) AND (fTargetBar <= DL_P_MAX)        // 目标压力在量程内
          AND (fHystBar >= 0.0) AND (fHystBar <= DL_HYST_MAX)     // 回差在量程内
          AND (fMinCycleS >= 0.0)                                 // 最小循环时间非负
          AND (fRecvM3 >= 0.0);                                   // 罐容积非负
xViable := xValid                                                // 有效为前提
            AND (_fHystClamp >= fHystNeedBar)                    // 回差不低于最小回差
            AND (fBufferM3 >= DL_BUF_MIN)                        // 缓冲容积达标
            AND (fLoadBar > DL_EPS);                             // 加载点须为正压
FC_DL_AirCompLoadUnloadHystCalc := xValid;                        // 返回码：TRUE = 计算可信

END_FUNCTION

(* ---- FC_DL_AirCompSpecificPowerCalc.st ---- *)
(*
  Name: FC_DL_AirCompSpecificPowerCalc
  Category: DL_Process
  Version: 1.0.0
  Round: R90 / 2026-11-25
  开源溯源：clean-room 自研（族 压缩空气系统能效，ST 开源生态实测 0 命中，无外部代码引入）
  功能：1) 比功率按「单位容积流量的轴功率」计算：fSpecificKW = 轴功率[kW] / 自由排气量[m3/min]，
           量纲为 kW/(m3/min)，是空压系统能效的第一评价指标（越小越优）。
        2) 折算单位能耗 fSecPerM3 按 1 kW = 1 kJ/s 换算：1 m3/min = 60 m3/h，故
           kJ/m3 = kW/(m3/min) × (1 kJ/s / 1 kW) × (60 s/min) = 比功率 × 60，
           该输出用于与电价直接相乘做年运行成本估算，单位是 kJ/m3（等价 kWh/1000 m3 需再除 3600）。
        3) 能效等级 iEffClass 按比功率门槛分级：0 = 优（≤ DL_KLASS1）、1 = 良（≤ DL_KLASS2）、
           2 = 及格（≤ DL_KLASS3）、3 = 差（> DL_KLASS3）。等级门槛为螺杆机常见量级，
           由 VAR CONSTANT 统一组态，不写死在算式里。
  边界条件：1) 非有限值闸：两路实值入参统一过 NOT(x > -DL_BIG AND x < DL_BIG)，
           同时拦 NaN 与 Inf，命中即拦断实值通路（两个 REAL 输出强制 0.0、等级置 3）并置无效（R19）。
        2) 分母零闸：ABS(fFadM3min) > DL_EPS 才允许相除；排气量为 0 表示空压机停机或流量计失流，
           比功率在数学上发散，故判无效而不是输出一个大数。
        3) 负值闸：轴功率为负（四象限变频回馈）与排气量为负（流量计反向）均判无效；
           回馈工况不属于本件的评价范围，不得用绝对值混入能效统计。
        4) 饱和钳制：比功率结果钳到 0 ~ DL_SP_MAX(200 kW/(m3/min))，避免极小排气量放大成无意义巨值；
           折算能耗同样钳到 0 ~ 12000 kJ/m3，与比功率上限按同一换算关系对齐（×60）。
        5) 量纲不一致的加法一律禁止：本件只有乘除，无跨量纲相加，等级判定只比较同量纲比功率。
  量纲自证：fSpecificKW = kW / (m3/min) = kW·min/m3 = kJ/m3 的 1/60（因 1 kW = 1 kJ/s）；
           fSecPerM3 = kW/(m3/min) × 60 (s/min) = kJ/m3，其中 60 为 [s/min] 时间换算因子；
           两输出量纲一致（同为 kJ/m3 的等价表述），等级门槛与 fSpecificKW 同量纲。
*)

FUNCTION FC_DL_AirCompSpecificPowerCalc : BOOL
VAR_INPUT
    fShaftKW      : REAL;   // 空压机轴功率 [kW] / Compressor shaft power [kW]
    fFadM3min     : REAL;   // 自由排气量 FAD [m3/min] / Free air delivery [m3/min]
END_VAR
VAR_OUTPUT
    fSpecificKW   : REAL;   // 比功率 [kW/(m3/min)] / Specific power [kW/(m3/min)]
    fSecPerM3     : REAL;   // 折算单位能耗 [kJ/m3] / Converted specific energy [kJ/m3]
    iEffClass     : INT;    // 能效等级 0..3（0 最优）[-] / Efficiency class 0..3, 0 best [-]
    xValid        : BOOL;   // 计算有效标志 [bool] / Calculation valid flag [bool]
END_VAR
VAR
    _fSpecRaw     : REAL;   // 未饱和的原始比功率 [kW/(m3/min)] / Raw specific power [kW/(m3/min)]
    _fSpecClamp   : REAL;   // 饱和钳制后的比功率 [kW/(m3/min)] / Clamped specific power [kW/(m3/min)]
END_VAR
VAR CONSTANT
    DL_EPS        : REAL := 1.0E-9;    // 分母零闸阈值 [-] / Division-zero gate threshold [-]
    DL_BIG        : REAL := 1.0E12;    // 非有限值闸量级上限 [-] / Finiteness gate magnitude [-]
    DL_S_PER_MIN  : REAL := 60.0;      // min → s 换算因子 [s/min] / Minute to second factor [s/min]
    DL_SP_MAX     : REAL := 200.0;     // 比功率饱和上限 [kW/(m3/min)] / Specific power saturation ceiling
    DL_KLASS1     : REAL := 5.0;       // 一级能效比功率门槛 [kW/(m3/min)] / Class-1 efficiency threshold
    DL_KLASS2     : REAL := 6.5;       // 二级能效比功率门槛 [kW/(m3/min)] / Class-2 efficiency threshold
    DL_KLASS3     : REAL := 8.5;       // 三级能效比功率门槛 [kW/(m3/min)] / Class-3 efficiency threshold
END_VAR

(* —— 段 1：非有限值闸（R19：闸断实值通路，NaN 不得进入除法） —— *)
IF NOT (fShaftKW > -DL_BIG AND fShaftKW < DL_BIG)
   OR NOT (fFadM3min > -DL_BIG AND fFadM3min < DL_BIG) THEN
    fSpecificKW := 0.0;                     // 输出强制 0.0 / Output forced to zero
    fSecPerM3 := 0.0;                       // 折算能耗强制 0.0 / Converted energy forced to zero
    iEffClass := 3;                         // 等级置最差档，不给误导性「优」/ Worst class only
    xValid := FALSE;                        // 有效位清零 / Validity cleared
    FC_DL_AirCompSpecificPowerCalc := FALSE;   // 返回码同源 / Return mirrors validity
    RETURN;                                 // 立即退出 / Immediate exit
END_IF

(* —— 段 2：组态与零闸（R4：分母先过 ABS 闸；负功率/负流量同属故障） —— *)
IF (ABS(fFadM3min) <= DL_EPS) OR (fShaftKW < 0.0) OR (fFadM3min < 0.0) THEN
    fSpecificKW := 0.0;                     // 输出强制 0.0 / Output forced to zero
    fSecPerM3 := 0.0;                       // 折算能耗强制 0.0 / Converted energy forced to zero
    iEffClass := 3;                         // 等级置最差档 / Worst class only
    xValid := FALSE;                        // 判无效 / Invalid
    FC_DL_AirCompSpecificPowerCalc := FALSE;   // 返回码同步 / Return synchronised
    RETURN;                                 // 提前退出 / Early exit
END_IF

(* —— 段 3：主算式（R22 方向自核：轴功率为分子、排气量为分母，不可取倒数） —— *)
_fSpecRaw := fShaftKW / fFadM3min;                          // 比功率 [kW/(m3/min)]
_fSpecClamp := LIMIT(0.0, _fSpecRaw, DL_SP_MAX);            // 饱和钳 0..200

(* —— 段 4：能效等级分级（IF/ELSIF 单链，iEffClass 只在此处赋值一次） —— *)
IF _fSpecClamp <= DL_KLASS1 THEN
    iEffClass := 0;                         // 一级能效（优）/ Class 1, best
ELSIF _fSpecClamp <= DL_KLASS2 THEN
    iEffClass := 1;                         // 二级能效（良）/ Class 2, good
ELSIF _fSpecClamp <= DL_KLASS3 THEN
    iEffClass := 2;                         // 三级能效（及格）/ Class 3, acceptable
ELSE
    iEffClass := 3;                         // 低于三级（差）/ Below class 3, poor
END_IF

(* —— 段 5：输出单点写盘（折算能耗与比功率同一基准，换算因子 60 s/min） —— *)
fSpecificKW := _fSpecClamp;                                 // 比功率出口 [kW/(m3/min)]
fSecPerM3 := _fSpecClamp * DL_S_PER_MIN;                    // 折算单位能耗 [kJ/m3]
xValid := (fShaftKW >= 0.0) AND (fFadM3min > DL_EPS);       // 有效位单点聚合
FC_DL_AirCompSpecificPowerCalc := xValid;                   // 返回码：TRUE = 计算可信

END_FUNCTION

(* ---- FC_DL_AirDewPointCalc.st ---- *)
(*
  Name: FC_DL_AirDewPointCalc
  Category: DL_Process
  Version: 1.0.0
  Round: R90 / 2026-11-25
  开源溯源：clean-room 自研（族 压缩空气系统能效，ST 开源生态实测 0 命中，无外部代码引入）
  功能：1) 压力露点 → 常压露点换算。物理口径：露点由「水蒸气分压」唯一确定，而分压等于
           摩尔分数乘总压。压缩空气从工作压力膨胀到大气压时摩尔分数不变、总压下降，
           故分压按 P_atm / P_abs 等比缩小，再由缩小后的分压反解露点即为常压露点。
           逐步为：Magnus 正解求工作压力下的饱和分压 → 按总压比缩小 → Magnus 反解温度。
        2) 含水量按理想气体状态方程在「压力露点温度」下计算：
           ρ[g/m3] = 1000 · p_v[Pa] / (R_v · T[K])，R_v = 461.5 J/(kg·K) 为水蒸气气体常数，
           合并常数后为 ρ = 2.1667 · p_v[Pa] / T[K]，表示工作压力下每立方米压缩空气的饱和含水量。
  边界条件：1) 非有限值闸：两路实值入参统一过 NOT(x > -DL_BIG AND x < DL_BIG)，
           同时拦 NaN 与 Inf，命中即拦断实值通路（两个 REAL 输出强制 0.0）并置无效（R19）。
        2) Magnus 分母零闸：DL_MAG_C + fPdpC 必须 ABS > DL_EPS，否则正解分母发散；
           反解分母 DL_MAG_B − L 同样必须 ABS > DL_EPS，否则常压露点发散。
        3) 开尔文偏移零闸：fPdpC + 273.15 > DL_EPS，否则含水量式温度分母为 0。
        4) 绝对值分母零闸：工作绝压 fWorkBar + DL_P_ATM_BAR 必须 ABS > DL_EPS（真空工况拦截）。
        5) 量程校验：压力露点 −90 ~ 100 °C（覆盖吸附式干燥机 −70 °C 到无油机高温工况），
           工作表压 0 ~ 100 bar；越域钳到边界算参考值但置无效。
        6) 饱和钳制：含水量钳 0 ~ 1000 g/m3，常压露点钳 −100 ~ 100 °C，防极端输入溢出。
  量纲自证：p_v = hPa × EXP([-]) = hPa，EXP 的自变量 (B·t)/(C+t) 中 (1/°C·°C) = 无因次；
           p_v_atm / p_v = (bar/bar) = 无因次，故分压换算不改变量纲；
           ADP 反解式 C·L/(B − L)：L = LN(hPa/hPa) 无因次，故结果为 °C；
           含水量 = 1000 [g/kg] × Pa / (J/(kg·K) × K) = g/m3，量纲闭合。
*)

FUNCTION FC_DL_AirDewPointCalc : BOOL
VAR_INPUT
    fPdpC         : REAL;   // 压力露点 [°C] / Pressure dew point [°C]
    fWorkBar      : REAL;   // 工作表压 [bar] / Working gauge pressure [bar]
END_VAR
VAR_OUTPUT
    fAdpC         : REAL;   // 常压露点 [°C] / Atmospheric dew point [°C]
    fMoistGm3     : REAL;   // 工作压力下饱和含水量 [g/m3] / Saturated moisture content [g/m3]
    xValid        : BOOL;   // 计算有效标志 [bool] / Calculation valid flag [bool]
END_VAR
VAR
    _fPdpClampC   : REAL;   // 钳制后的压力露点 [°C] / Clamped pressure dew point [°C]
    _fPAbsBar     : REAL;   // 工作绝对压力 [bar] / Working absolute pressure [bar]
    _fPvHpa       : REAL;   // 工作压力下饱和水蒸气分压 [hPa] / Saturation vapour pressure [hPa]
    _fPvAtmHpa    : REAL;   // 膨胀到常压后的水蒸气分压 [hPa] / Vapour pressure after expansion [hPa]
    _fL           : REAL;   // Magnus 反解中间量 LN(p_v/6.112) [-] / Magnus inverse intermediate [-]
    _fAdpRawC     : REAL;   // 未饱和的常压露点 [°C] / Raw atmospheric dew point [°C]
    _fMoistRaw    : REAL;   // 未饱和的含水量 [g/m3] / Raw moisture content [g/m3]
    _bDenOk       : BOOL;   // 三个分母合法性聚合 [bool] / Three denominator validity aggregate [bool]
END_VAR
VAR CONSTANT
    DL_EPS        : REAL := 1.0E-9;    // 分母零闸阈值 [-] / Division-zero gate threshold [-]
    DL_BIG        : REAL := 1.0E12;    // 非有限值闸量级上限 [-] / Finiteness gate magnitude [-]
    DL_MAG_A      : REAL := 6.112;     // Magnus 系数 A（0 °C 饱和压）[hPa] / Magnus coefficient A [hPa]
    DL_MAG_B      : REAL := 17.62;     // Magnus 系数 B [-]/ Magnus coefficient B [-]
    DL_MAG_C      : REAL := 243.12;    // Magnus 系数 C [°C] / Magnus coefficient C [°C]
    DL_K0         : REAL := 273.15;    // 摄氏转开尔文偏移 [K] / Celsius to Kelvin offset [K]
    DL_P_ATM_BAR  : REAL := 1.01325;   // 标准大气压 [bar] / Standard atmospheric pressure [bar]
    DL_RHOV_K     : REAL := 2.1667;    // 水蒸气密度合并常数 [g·K/(m3·Pa)] / Vapour density constant
    DL_PDP_LO_C   : REAL := -90.0;     // 压力露点量程下限 [°C] / Pressure dew point range low [°C]
    DL_PDP_HI_C   : REAL := 100.0;     // 压力露点量程上限 [°C] / Pressure dew point range high [°C]
    DL_P_LO_BAR   : REAL := 0.0;       // 工作表压量程下限 [bar] / Gauge pressure range low [bar]
    DL_P_HI_BAR   : REAL := 100.0;     // 工作表压量程上限 [bar] / Gauge pressure range high [bar]
    DL_ADP_LO_C   : REAL := -100.0;    // 常压露点饱和下限 [°C] / Atmospheric dew point low [°C]
    DL_ADP_HI_C   : REAL := 100.0;     // 常压露点饱和上限 [°C] / Atmospheric dew point high [°C]
    DL_MOIST_MAX  : REAL := 1000.0;    // 含水量饱和上限 [g/m3] / Moisture saturation ceiling [g/m3]
END_VAR

(* —— 段 1：非有限值闸（R19：闸断实值通路，NaN 不得进 EXP/LN） —— *)
IF NOT (fPdpC > -DL_BIG AND fPdpC < DL_BIG)
   OR NOT (fWorkBar > -DL_BIG AND fWorkBar < DL_BIG) THEN
    fAdpC := 0.0;                           // 输出强制 0.0 / Output forced to zero
    fMoistGm3 := 0.0;                       // 含水量强制 0.0 / Moisture forced to zero
    xValid := FALSE;                        // 有效位清零 / Validity cleared
    FC_DL_AirDewPointCalc := FALSE;         // 返回码同源 / Return mirrors validity
    RETURN;                                 // 立即退出 / Immediate exit
END_IF

(* —— 段 2：分母零闸（R4：Magnus 分母、绝对压分母、开尔文分母三处逐一验证） —— *)
_fPAbsBar := fWorkBar + DL_P_ATM_BAR;       // 工作绝压 [bar]
_bDenOk := (ABS(DL_MAG_C + fPdpC) > DL_EPS)                       // Magnus 正解分母
           AND (_fPAbsBar > DL_EPS)                               // 绝对压分母（真空拦截）
           AND ((fPdpC + DL_K0) > DL_EPS);                        // 含水量开尔文分母
IF NOT _bDenOk THEN
    fAdpC := 0.0;                           // 输出强制 0.0 / Output forced to zero
    fMoistGm3 := 0.0;                       // 含水量强制 0.0 / Moisture forced to zero
    xValid := FALSE;                        // 判无效 / Invalid
    FC_DL_AirDewPointCalc := FALSE;         // 返回码同步 / Return synchronised
    RETURN;                                 // 提前退出 / Early exit
END_IF

(* —— 段 3：量程钳制（越域钳边界算参考值，段 6 判无效） —— *)
_fPdpClampC := LIMIT(DL_PDP_LO_C, fPdpC, DL_PDP_HI_C);            // 压力露点钳 −90..100 [°C]

(* —— 段 4：Magnus 正解求分压（R22 方向自核：露点升高→分压升高，指数为正） —— *)
_fPvHpa := DL_MAG_A * EXP(DL_MAG_B * _fPdpClampC / (DL_MAG_C + _fPdpClampC));   // [hPa]
_fPvAtmHpa := _fPvHpa * DL_P_ATM_BAR / _fPAbsBar;                                // 膨胀后分压 [hPa]

(* —— 段 5：Magnus 反解常压露点（分母 B − L 已闸，L >= B 时判无效） —— *)
_fL := LN(MAX(DL_EPS, _fPvAtmHpa / DL_MAG_A));                     // LN(p_v/A) [-]
IF ABS(DL_MAG_B - _fL) > DL_EPS THEN
    _fAdpRawC := DL_MAG_C * _fL / (DL_MAG_B - _fL);                // 常压露点 [°C]
ELSE
    _fAdpRawC := DL_ADP_LO_C;                                      // 分母发散：退下限哨兵值
END_IF

(* —— 段 6：含水量（工作压力、压力露点温度下的饱和含水量） —— *)
_fMoistRaw := DL_RHOV_K * (_fPvHpa * 100.0) / (_fPdpClampC + DL_K0);   // ρ [g/m3]

(* —— 段 7：有效位单点聚合（量程 + 反解分母合法） —— *)
xValid := (fPdpC >= DL_PDP_LO_C) AND (fPdpC <= DL_PDP_HI_C)        // 压力露点在量程内
          AND (fWorkBar >= DL_P_LO_BAR) AND (fWorkBar <= DL_P_HI_BAR)   // 工作压力在量程内
          AND (ABS(DL_MAG_B - _fL) > DL_EPS);                      // 反解分母不发散

(* —— 段 8：输出单点写盘（饱和钳制） —— *)
fAdpC := LIMIT(DL_ADP_LO_C, _fAdpRawC, DL_ADP_HI_C);               // 常压露点 [°C]
fMoistGm3 := LIMIT(0.0, _fMoistRaw, DL_MOIST_MAX);                 // 含水量 [g/m3]
FC_DL_AirDewPointCalc := xValid;                                   // 返回码：TRUE = 计算可信

END_FUNCTION

(* ---- FC_DL_AirDryerPurgeLossCalc.st ---- *)
(*
  Name: FC_DL_AirDryerPurgeLossCalc
  Category: DL_Process
  Version: 1.0.0
  Round: R90 / 2026-11-25
  开源溯源：clean-room 自研（族 压缩空气系统能效，ST 开源生态实测 0 命中，无外部代码引入）
  功能：1) 吸附式干燥机再生耗气量按「额定处理流量 × 再生耗气率」计算：
           fLossM3min = fRatedFlowM3min × fPurgePct / 100。再生耗气是无谓损耗，
           它同时意味着上游空压机要多产这部分气，故必须计入系统能耗。
        2) 年运行成本按「损耗气量 → 等效电耗 → 电费」三段折算：
             等效比功率 = 额定轴功率 / 额定处理流量，量纲 kW/(m3/min)；
             年电耗[kWh] = 损耗气量[m3/min] × 比功率[kW/(m3/min)] × 年运行小时[h]；
             年成本 = 年电耗 × 电价。注意比功率已按「每分钟气量」定义，
             故乘年小时数即可，不得再乘 60 做时间换算（这是本件最容易写错的一处方向问题）。
  边界条件：1) 非有限值闸：五路实值入参统一过 NOT(x > -DL_BIG AND x < DL_BIG)，
           同时拦 NaN 与 Inf，命中即拦断实值通路（两个 REAL 输出强制 0.0）并置无效（R19）。
        2) 分母零闸：ABS(fRatedFlowM3min) > DL_EPS 才能得到比功率，
           额定流量为 0 表示铭牌未录入，判无效而不是输出无意义成本。
        3) 负值闸：额定流量、再生耗气率、年运行小时、电价、额定功率任一为负判无效
           （再生耗气率为负会得出「负成本」，属组态错误，不取绝对值掩盖）。
        4) 量程校验：再生耗气率必须落在 0 ~ 100 %（超过 100 % 意味着再生耗气大于处理量，
           干燥机不可能工作），年运行小时钳 0 ~ 8760 h，电价钳 0 ~ DL_PRICE_MAX。
        5) 饱和钳制：耗气量钳 0 ~ DL_LOSS_MAX，年成本钳 0 ~ DL_COST_MAX，防溢出。
  量纲自证：fLossM3min = (m3/min) × (%/100) = m3/min；
           比功率 = kW / (m3/min) = kW·min/m3；
           年电耗 = (m3/min) × (kW·min/m3) × h = kW·h，量纲闭合（min 与 min 对消）；
           年成本 = kWh × (货币/kWh) = 货币，三项内部量纲一致，未出现 kW/kW 去加温度的混算。
*)

FUNCTION FC_DL_AirDryerPurgeLossCalc : BOOL
VAR_INPUT
    fRatedFlowM3min : REAL;   // 干燥机额定处理流量 [m3/min] / Dryer rated flow [m3/min]
    fPurgePct       : REAL;   // 再生耗气率 [%] / Regeneration purge ratio [%]
    fHoursYear      : REAL;   // 年运行小时数 [h] / Annual operating hours [h]
    fPricePerKWh    : REAL;   // 电价 [货币/kWh] / Electricity price [currency/kWh]
    fRatedKW        : REAL;   // 空压机额定轴功率 [kW] / Compressor rated shaft power [kW]
END_VAR
VAR_OUTPUT
    fLossM3min      : REAL;   // 再生耗气量 [m3/min] / Regeneration purge loss [m3/min]
    fSpecKW         : REAL;   // 等效比功率 [kW/(m3/min)] / Equivalent specific power [kW/(m3/min)]
    fCostYear       : REAL;   // 年运行成本 [货币] / Annual operating cost [currency]
    xValid          : BOOL;   // 计算有效标志 [bool] / Calculation valid flag [bool]
END_VAR
VAR
    _fSpecRaw       : REAL;   // 未饱和的等效比功率 [kW/(m3/min)] / Raw specific power
    _fPurgeRatio    : REAL;   // 归一化再生耗气率 [-] / Normalized purge ratio [-]
    _fLossRaw       : REAL;   // 未饱和的耗气量 [m3/min] / Raw purge loss [m3/min]
    _fHoursClamp    : REAL;   // 钳制后的年运行小时 [h] / Clamped annual hours [h]
    _fCostRaw       : REAL;   // 未饱和的年成本 [货币] / Raw annual cost [currency]
END_VAR
VAR CONSTANT
    DL_EPS          : REAL := 1.0E-9;    // 分母零闸阈值 [-] / Division-zero gate threshold [-]
    DL_BIG          : REAL := 1.0E12;    // 非有限值闸量级上限 [-] / Finiteness gate magnitude [-]
    DL_PCT          : REAL := 100.0;     // 百分比换算因子 [%] / Percent conversion factor [%]
    DL_HOURS_YEAR   : REAL := 8760.0;    // 全年小时数上限 [h] / Hours per year upper bound [h]
    DL_PRICE_MAX    : REAL := 100.0;     // 电价量程上限 [货币/kWh] / Electricity price ceiling
    DL_LOSS_MAX     : REAL := 10000.0;   // 耗气量饱和上限 [m3/min] / Purge loss saturation ceiling [m3/min]
    DL_COST_MAX     : REAL := 1.0E9;     // 年成本饱和上限 [货币] / Annual cost saturation ceiling
END_VAR

(* —— 段 1：非有限值闸（R19：五路入参全覆盖，拦 NaN 与 Inf） —— *)
IF NOT (fRatedFlowM3min > -DL_BIG AND fRatedFlowM3min < DL_BIG)
   OR NOT (fPurgePct > -DL_BIG AND fPurgePct < DL_BIG)
   OR NOT (fHoursYear > -DL_BIG AND fHoursYear < DL_BIG)
   OR NOT (fPricePerKWh > -DL_BIG AND fPricePerKWh < DL_BIG)
   OR NOT (fRatedKW > -DL_BIG AND fRatedKW < DL_BIG) THEN
    fLossM3min := 0.0;                      // 输出强制 0.0 / Output forced to zero
    fSpecKW := 0.0;                         // 比功率强制 0.0 / Specific power forced to zero
    fCostYear := 0.0;                       // 成本强制 0.0 / Cost forced to zero
    xValid := FALSE;                        // 有效位清零 / Validity cleared
    FC_DL_AirDryerPurgeLossCalc := FALSE;   // 返回码同源 / Return mirrors validity
    RETURN;                                 // 立即退出 / Immediate exit
END_IF

(* —— 段 2：分母零闸（R4：额定流量是比功率的分母，必须先过 ABS 闸） —— *)
IF ABS(fRatedFlowM3min) <= DL_EPS THEN
    fLossM3min := 0.0;                      // 输出强制 0.0 / Output forced to zero
    fSpecKW := 0.0;                         // 比功率强制 0.0 / Specific power forced to zero
    fCostYear := 0.0;                       // 成本强制 0.0 / Cost forced to zero
    xValid := FALSE;                        // 判无效 / Invalid
    FC_DL_AirDryerPurgeLossCalc := FALSE;   // 返回码同步 / Return synchronised
    RETURN;                                 // 提前退出 / Early exit
END_IF

(* —— 段 3：负值闸（负耗气率会得出负成本，属组态错误） —— *)
IF (fRatedFlowM3min < 0.0) OR (fPurgePct < 0.0) OR (fHoursYear < 0.0)
   OR (fPricePerKWh < 0.0) OR (fRatedKW < 0.0) THEN
    fLossM3min := 0.0;                      // 输出强制 0.0 / Output forced to zero
    fSpecKW := 0.0;                         // 比功率强制 0.0 / Specific power forced to zero
    fCostYear := 0.0;                       // 成本强制 0.0 / Cost forced to zero
    xValid := FALSE;                        // 判无效 / Invalid
    FC_DL_AirDryerPurgeLossCalc := FALSE;   // 返回码同步 / Return synchronised
    RETURN;                                 // 提前退出 / Early exit
END_IF

(* —— 段 4：等效比功率（R22 方向自核：额定功率在分子，额定流量在分母） —— *)
_fSpecRaw := fRatedKW / fRatedFlowM3min;                          // [kW/(m3/min)]

(* —— 段 5：再生耗气量与年成本（比功率已按每分钟定义，故不再乘 60） —— *)
_fPurgeRatio := fPurgePct / DL_PCT;                               // 归一化 [-]
_fLossRaw := fRatedFlowM3min * _fPurgeRatio;                      // 耗气量 [m3/min]
_fHoursClamp := LIMIT(0.0, fHoursYear, DL_HOURS_YEAR);            // 年小时钳制 [h]
_fCostRaw := _fLossRaw * _fSpecRaw * _fHoursClamp * fPricePerKWh; // 年成本 [货币]

(* —— 段 6：输出单点写盘（饱和钳制） —— *)
fSpecKW := LIMIT(0.0, _fSpecRaw, DL_BIG);                         // 比功率 [kW/(m3/min)]
fLossM3min := LIMIT(0.0, _fLossRaw, DL_LOSS_MAX);                 // 耗气量 [m3/min]
fCostYear := LIMIT(0.0, _fCostRaw, DL_COST_MAX);                  // 年成本 [货币]

(* —— 段 7：有效位单点聚合（耗气率窄闸 + 电价量程） —— *)
xValid := (fRatedFlowM3min > DL_EPS)                              // 额定流量为正
          AND (fPurgePct <= DL_PCT)                               // 耗气率不超 100 %
          AND (fHoursYear <= DL_HOURS_YEAR)                       // 年小时不超 8760
          AND (fPricePerKWh <= DL_PRICE_MAX)                      // 电价在量程内
          AND (fRatedKW >= 0.0);                                  // 额定功率非负
FC_DL_AirDryerPurgeLossCalc := xValid;                            // 返回码：TRUE = 计算可信

END_FUNCTION

(* ---- FC_DL_AirLeakRateCalc.st ---- *)
(*
  Name: FC_DL_AirLeakRateCalc
  Category: DL_Process
  Version: 1.0.0
  Round: R90 / 2026-11-25
  开源溯源：clean-room 自研（族 压缩空气系统能效，ST 开源生态实测 0 命中，无外部代码引入）
  功能：1) 停机压降法测泄漏流量：全厂停机（无生产用气）后记录储气罐从 P1 降到 P2 的时长，
           罐内减少的「常压自由空气容积」= 罐容积 × (P1 − P2) / 大气压，
           折算到每分钟即泄漏流量：fLeakM3min = V · (P1 − P2) / P_atm · 60 / t。
           泄漏流量的方向是「从罐内流向大气」，故压降为 P1 − P2（前减后），不可反写。
        2) 泄漏占比：fLeakPct = 泄漏流量 / 平均用气需求 × 100，
           分母是生产期实测平均需求（同量纲 m3/min），用来判断泄漏占总耗气的份额；
           该口径对应「改造泄漏可节省的最大气量比例」，不是压缩机能耗占比。
  边界条件：1) 非有限值闸：五路实值入参统一过 NOT(x > -DL_BIG AND x < DL_BIG)，
           同时拦 NaN 与 Inf，命中即拦断实值通路（两个 REAL 输出强制 0.0）并置无效（R19）。
        2) 分母零闸：ABS(fTimeS) > DL_EPS 与 ABS(fAvgDemandM3min) > DL_EPS 都必须通过；
           测量时长为 0 则泄漏流量发散，平均需求为 0 则占比发散（无生产工况无法归一）。
        3) 分母零闸补充：ABS(DL_P_ATM_BAR) 为常量不可能为零，但仍以常量直接使用（编译期确定），
           不引入运行期除法风险。
        4) 压降方向闸：fP1Bar 必须 > fP2Bar，否则压降为负（记录顺序颠倒或罐被充气），判无效；
           压降为 0 属合法但无信息，输出 0 且判无效（无压降无法算出泄漏）。
        5) 负值闸：罐容积、压力、时长、需求任一为负判无效（不取绝对值掩盖反向）。
        6) 饱和钳制：泄漏流量钳 0 ~ DL_LEAK_MAX(10000 m3/min)，占比钳 0 ~ 100 %，
           防极短测量时长把泄漏值放大到无意义量级。
  量纲自证：V·ΔP/P_atm = m3 × bar / bar = m3；× 60 [s/min] / t[s] → m3/min；
           fLeakPct = (m3/min) / (m3/min) × 100 = 无因次百分数 [%]，分母与分子同量纲。
*)

FUNCTION FC_DL_AirLeakRateCalc : BOOL
VAR_INPUT
    fTankM3          : REAL;   // 储气罐有效容积 [m3] / Effective receiver volume [m3]
    fP1Bar           : REAL;   // 起始罐压 [bar] / Initial receiver pressure [bar]
    fP2Bar           : REAL;   // 结束罐压 [bar] / Final receiver pressure [bar]
    fTimeS           : REAL;   // 测量时长 [s] / Measurement duration [s]
    fAvgDemandM3min  : REAL;   // 生产期平均用气需求 [m3/min] / Average production air demand [m3/min]
END_VAR
VAR_OUTPUT
    fLeakM3min       : REAL;   // 泄漏流量 [m3/min] / Leakage flow [m3/min]
    fLeakPct         : REAL;   // 泄漏占平均需求比例 [%] / Leakage share of average demand [%]
    xValid           : BOOL;   // 计算有效标志 [bool] / Calculation valid flag [bool]
END_VAR
VAR
    _fDropBar        : REAL;   // 测量期间压降 [bar] / Pressure drop during test [bar]
    _fFreeVolumeM3   : REAL;   // 压降对应的常压自由空气容积 [m3] / Free air volume from drop [m3]
    _fLeakRawM3min   : REAL;   // 未饱和的泄漏流量 [m3/min] / Raw leakage flow [m3/min]
    _fLeakPctRaw     : REAL;   // 未饱和的泄漏占比 [%] / Raw leakage share [%]
END_VAR
VAR CONSTANT
    DL_EPS           : REAL := 1.0E-9;    // 分母零闸阈值 [-] / Division-zero gate threshold [-]
    DL_BIG           : REAL := 1.0E12;    // 非有限值闸量级上限 [-] / Finiteness gate magnitude [-]
    DL_P_ATM_BAR     : REAL := 1.01325;   // 标准大气压 [bar] / Standard atmospheric pressure [bar]
    DL_S_PER_MIN     : REAL := 60.0;      // min → s 换算因子 [s/min] / Minute to second factor [s/min]
    DL_PCT           : REAL := 100.0;     // 百分比换算因子 [%] / Percent conversion factor [%]
    DL_LEAK_MAX      : REAL := 10000.0;   // 泄漏流量饱和上限 [m3/min] / Leakage saturation ceiling [m3/min]
    DL_DROP_MIN      : REAL := 1.0E-6;    // 压降有效下限 [bar] / Minimum meaningful pressure drop [bar]
END_VAR

(* —— 段 1：非有限值闸（R19：五路入参全覆盖，拦 NaN 与 Inf） —— *)
IF NOT (fTankM3 > -DL_BIG AND fTankM3 < DL_BIG)
   OR NOT (fP1Bar > -DL_BIG AND fP1Bar < DL_BIG)
   OR NOT (fP2Bar > -DL_BIG AND fP2Bar < DL_BIG)
   OR NOT (fTimeS > -DL_BIG AND fTimeS < DL_BIG)
   OR NOT (fAvgDemandM3min > -DL_BIG AND fAvgDemandM3min < DL_BIG) THEN
    fLeakM3min := 0.0;                      // 输出强制 0.0 / Output forced to zero
    fLeakPct := 0.0;                        // 占比强制 0.0 / Share forced to zero
    xValid := FALSE;                        // 有效位清零 / Validity cleared
    FC_DL_AirLeakRateCalc := FALSE;         // 返回码同源 / Return mirrors validity
    RETURN;                                 // 立即退出 / Immediate exit
END_IF

(* —— 段 2：分母零闸（R4：测量时长与平均需求两个分母逐一验证） —— *)
IF (ABS(fTimeS) <= DL_EPS) OR (ABS(fAvgDemandM3min) <= DL_EPS) THEN
    fLeakM3min := 0.0;                      // 输出强制 0.0 / Output forced to zero
    fLeakPct := 0.0;                        // 占比强制 0.0 / Share forced to zero
    xValid := FALSE;                        // 判无效 / Invalid
    FC_DL_AirLeakRateCalc := FALSE;         // 返回码同步 / Return synchronised
    RETURN;                                 // 提前退出 / Early exit
END_IF

(* —— 段 3：负值闸与压降方向闸（R22：压降是前减后，方向颠倒即判无效） —— *)
_fDropBar := fP1Bar - fP2Bar;               // 测量期间压降（前 − 后）[bar]
IF (fTankM3 < 0.0) OR (fTimeS < 0.0) OR (fAvgDemandM3min < 0.0) OR (_fDropBar < 0.0) THEN
    fLeakM3min := 0.0;                      // 输出强制 0.0 / Output forced to zero
    fLeakPct := 0.0;                        // 占比强制 0.0 / Share forced to zero
    xValid := FALSE;                        // 判无效 / Invalid
    FC_DL_AirLeakRateCalc := FALSE;         // 返回码同步 / Return synchronised
    RETURN;                                 // 提前退出 / Early exit
END_IF

(* —— 段 4：泄漏流量主算式（压降 → 常压容积 → 每分钟） —— *)
_fFreeVolumeM3 := fTankM3 * _fDropBar / DL_P_ATM_BAR;             // 常压自由空气容积 [m3]
_fLeakRawM3min := _fFreeVolumeM3 * DL_S_PER_MIN / fTimeS;         // 泄漏流量 [m3/min]

(* —— 段 5：泄漏占比（分母为平均需求，同量纲归一化） —— *)
_fLeakPctRaw := _fLeakRawM3min / fAvgDemandM3min * DL_PCT;        // 占比 [%]

(* —— 段 6：有效位单点聚合（压降必须有效，无压降无法算泄漏） —— *)
xValid := (_fDropBar > DL_DROP_MIN)                               // 压降有效
          AND (fTankM3 > 0.0)                                     // 罐容积为正
          AND (fTimeS > DL_EPS)                                   // 测量时长为正
          AND (fAvgDemandM3min > DL_EPS);                         // 平均需求为正（占比可归一）

(* —— 段 7：输出单点写盘（饱和钳制） —— *)
fLeakM3min := LIMIT(0.0, _fLeakRawM3min, DL_LEAK_MAX);            // 泄漏流量 [m3/min]
fLeakPct := LIMIT(0.0, _fLeakPctRaw, DL_PCT);                     // 泄漏占比钳 0..100 [%]
FC_DL_AirLeakRateCalc := xValid;                                  // 返回码：TRUE = 计算可信

END_FUNCTION

(* ---- FC_DL_AirNozzleConsumptionCalc.st ---- *)
(*
  Name: FC_DL_AirNozzleConsumptionCalc
  Category: DL_Process
  Version: 1.0.0
  Round: R90 / 2026-11-25
  开源溯源：clean-room 自研（族 压缩空气系统能效，ST 开源生态实测 0 命中，无外部代码引入）
  功能：1) 单喷嘴耗气量按喷管临界（声速）流模型计算：当供气压力与背压之比超过临界比时，
           喉部达到声速，质量流量只取决于上游绝对压力而与背压无关，即
             m_dot = Cd · A · P_abs · sqrt(k/(R·T)) · (2/(k+1))^((k+1)/(2(k-1)))
           其中 k = 1.4、R = 287 J/(kg·K)、T = 293.15 K，合并为一个常数 DL_MDOT_K，
           故 m_dot = Cd · A · P_abs · DL_MDOT_K [kg/s]。
        2) 质量流量折算为常压自由空气体积流量：除以常压密度 DL_RHO_N(1.2046 kg/m3)，
           再乘 60 得 m3/min，即 fPerNozzleM3min。
        3) 总耗气量 = 单喷嘴耗气量 × 喷嘴数量 × 同时使用率 / 100。使用率是「同时吹气的比例」，
           按百分比归一化后乘入，方向为放大系数（使用率越高总耗气越大）。
  边界条件：1) 非有限值闸：三路实值入参统一过 NOT(x > -DL_BIG AND x < DL_BIG)，
           同时拦 NaN 与 Inf，命中即拦断实值通路（两个 REAL 输出强制 0.0）并置无效（R19）。
        2) 分母零闸：本件除数均为常量（DL_RHO_N、100.0），无常量零风险；
           但喷嘴口径与绝对压力的乘积必须为正，故对 fOrificeMm 做 DL_D_MIN_MM(0.1 mm) 下限钳制，
           防口径为 0 使耗气量恒为 0 而掩盖配置错误。
        3) 数量零闸：iCount < 0 判无效（负数量无物理意义）；iCount = 0 属合法（该支路无喷嘴），
           总耗气输出 0，不判无效。
        4) 使用率窄闸：fUsePct 必须落在 0 ~ 100 %，越域钳到边界并置无效；
           负使用率不取绝对值（会虚增耗气）。
        5) 饱和钳制：绝对压力按 DL_P_ABS_MAX(101 bar) 上限钳制，单喷嘴耗气钳 0 ~ 100 m3/min，
           总耗气钳 0 ~ 100000 m3/min，防数量与口径同时极端时溢出。
  量纲自证：A = m2，P_abs = Pa，DL_MDOT_K = kg/(s·m2·Pa)，故 m_dot = kg/s；
           除以 DL_RHO_N(kg/m3) → m3/s，乘 60 s/min → m3/min；
           总耗气 = (m3/min) × [-] × (%/100) = m3/min，百分比为无因次比例。
*)

FUNCTION FC_DL_AirNozzleConsumptionCalc : BOOL
VAR_INPUT
    fOrificeMm     : REAL;   // 喷嘴等效口径 [mm] / Nozzle equivalent orifice diameter [mm]
    fSupplyBar     : REAL;   // 供气表压 [bar] / Supply gauge pressure [bar]
    iCount         : INT;    // 喷嘴数量 [个] / Nozzle count [pcs]
    fUsePct        : REAL;   // 同时使用率 [%] / Simultaneous use ratio [%]
END_VAR
VAR_OUTPUT
    fPerNozzleM3min: REAL;   // 单喷嘴耗气量 [m3/min] / Consumption per nozzle [m3/min]
    fTotalM3min    : REAL;   // 总耗气量 [m3/min] / Total consumption [m3/min]
    fVelMps        : REAL;   // 喷嘴出口等效流速（观测用）[m/s] / Equivalent exit velocity [m/s]
    xValid         : BOOL;   // 计算有效标志 [bool] / Calculation valid flag [bool]
END_VAR
VAR
    _fDClampMm     : REAL;   // 钳制后的口径 [mm] / Clamped orifice diameter [mm]
    _fAreaM2       : REAL;   // 喷嘴截面积 [m2] / Nozzle cross-section area [m2]
    _fPAbsPa       : REAL;   // 供气绝对压力 [Pa] / Supply absolute pressure [Pa]
    _fMDotKgS      : REAL;   // 质量流量 [kg/s] / Mass flow rate [kg/s]
    _fPerRawM3min  : REAL;   // 未饱和的单喷嘴耗气量 [m3/min] / Raw per-nozzle consumption [m3/min]
    _fUseRatio     : REAL;   // 归一化使用率 [-] / Normalized use ratio [-]
    _fCountReal    : REAL;   // 数量的实数形态 [个] / Nozzle count as real [pcs]
    _fTotalRaw     : REAL;   // 未饱和的总耗气量 [m3/min] / Raw total consumption [m3/min]
END_VAR
VAR CONSTANT
    DL_EPS         : REAL := 1.0E-9;    // 分母零闸阈值 [-] / Division-zero gate threshold [-]
    DL_BIG         : REAL := 1.0E12;    // 非有限值闸量级上限 [-] / Finiteness gate magnitude [-]
    DL_PCT         : REAL := 100.0;     // 百分比换算因子 [%] / Percent conversion factor [%]
    DL_PI          : REAL := 3.14159265;   // 圆周率 [-] / Pi [-]
    DL_MM_PER_M    : REAL := 1000.0;    // m → mm 换算因子 [mm/m] / Metre to millimetre factor [mm/m]
    DL_S_PER_MIN   : REAL := 60.0;      // min → s 换算因子 [s/min] / Minute to second factor [s/min]
    DL_PA_PER_BAR  : REAL := 1.0E5;     // Pa → bar 换算因子 [Pa/bar] / Pascal to bar factor [Pa/bar]
    DL_P_ATM_BAR   : REAL := 1.01325;   // 标准大气压 [bar] / Standard atmospheric pressure [bar]
    DL_P_ABS_MAX   : REAL := 101.0;     // 绝对压力饱和上限 [bar] / Absolute pressure saturation ceiling [bar]
    DL_CD          : REAL := 0.65;      // 喷嘴流量系数 Cd [-] / Nozzle discharge coefficient Cd [-]
    DL_MDOT_K      : REAL := 2.362E-3;  // 临界流合并常数 [kg/(s·m2·Pa)] / Choked-flow lumped constant
    DL_RHO_N       : REAL := 1.2046;    // 常压 20 °C 空气密度 [kg/m3] / Air density at 20 degC 1 atm [kg/m3]
    DL_D_MIN_MM    : REAL := 0.10;      // 口径下限钳制值 [mm] / Orifice lower clamp [mm]
    DL_PER_MAX     : REAL := 100.0;     // 单喷嘴耗气饱和上限 [m3/min] / Per-nozzle saturation ceiling [m3/min]
    DL_TOT_MAX     : REAL := 100000.0;  // 总耗气饱和上限 [m3/min] / Total saturation ceiling [m3/min]
END_VAR

(* —— 段 1：非有限值闸（R19：三路实值入参全覆盖，拦 NaN 与 Inf） —— *)
IF NOT (fOrificeMm > -DL_BIG AND fOrificeMm < DL_BIG)
   OR NOT (fSupplyBar > -DL_BIG AND fSupplyBar < DL_BIG)
   OR NOT (fUsePct > -DL_BIG AND fUsePct < DL_BIG) THEN
    fPerNozzleM3min := 0.0;                 // 输出强制 0.0 / Output forced to zero
    fTotalM3min := 0.0;                     // 总耗气强制 0.0 / Total forced to zero
    fVelMps := 0.0;                         // 观测流速强制 0.0 / Velocity forced to zero
    xValid := FALSE;                        // 有效位清零 / Validity cleared
    FC_DL_AirNozzleConsumptionCalc := FALSE;   // 返回码同源 / Return mirrors validity
    RETURN;                                 // 立即退出 / Immediate exit
END_IF

(* —— 段 2：组态闸（口径为正、数量非负、供压非负） —— *)
IF (fOrificeMm <= DL_EPS) OR (iCount < 0) OR (fSupplyBar < 0.0) THEN
    fPerNozzleM3min := 0.0;                 // 输出强制 0.0 / Output forced to zero
    fTotalM3min := 0.0;                     // 总耗气强制 0.0 / Total forced to zero
    fVelMps := 0.0;                         // 观测流速强制 0.0 / Velocity forced to zero
    xValid := FALSE;                        // 判无效 / Invalid
    FC_DL_AirNozzleConsumptionCalc := FALSE;   // 返回码同步 / Return synchronised
    RETURN;                                 // 提前退出 / Early exit
END_IF

(* —— 段 3：几何与压力换算（口径下限钳制，绝对压上限钳制） —— *)
_fDClampMm := MAX(DL_D_MIN_MM, fOrificeMm);                        // 口径下限钳 [mm]
_fAreaM2 := DL_PI * (_fDClampMm / DL_MM_PER_M) * (_fDClampMm / DL_MM_PER_M) / 4.0;   // 截面积 [m2]
_fPAbsPa := LIMIT(0.0, fSupplyBar + DL_P_ATM_BAR, DL_P_ABS_MAX) * DL_PA_PER_BAR;      // 绝对压 [Pa]

(* —— 段 4：临界流质量流量（R22 方向自核：压力在分子，临界比已并入常数） —— *)
_fMDotKgS := DL_CD * _fAreaM2 * _fPAbsPa * DL_MDOT_K;              // 质量流量 [kg/s]

(* —— 段 5：质量流量 → 常压体积流量；再乘数量与使用率 —— *)
_fPerRawM3min := _fMDotKgS / DL_RHO_N * DL_S_PER_MIN;              // 单喷嘴耗气 [m3/min]
_fUseRatio := LIMIT(0.0, fUsePct, DL_PCT) / DL_PCT;                // 使用率归一 [-]
_fCountReal := INT_TO_REAL(iCount);                                // 数量实数化 [个]
_fTotalRaw := _fPerRawM3min * _fCountReal * _fUseRatio;            // 总耗气 [m3/min]

(* —— 段 6：输出单点写盘（饱和钳制，观测流速按单喷嘴流量反算等效出口流速） —— *)
fPerNozzleM3min := LIMIT(0.0, _fPerRawM3min, DL_PER_MAX);          // 单喷嘴耗气 [m3/min]
fTotalM3min := LIMIT(0.0, _fTotalRaw, DL_TOT_MAX);                 // 总耗气 [m3/min]
fVelMps := LIMIT(0.0, (fPerNozzleM3min / DL_S_PER_MIN) / _fAreaM2, DL_BIG);   // 等效流速 [m/s]

(* —— 段 7：有效位单点聚合（使用率不越域 + 口径与数量合法） —— *)
xValid := (fUsePct >= 0.0) AND (fUsePct <= DL_PCT)                 // 使用率在 0..100 %
          AND (fOrificeMm > DL_EPS)                                // 口径为正
          AND (iCount >= 0)                                        // 数量非负
          AND (fSupplyBar >= 0.0);                                 // 供压非负
FC_DL_AirNozzleConsumptionCalc := xValid;                          // 返回码：TRUE = 计算可信

END_FUNCTION

(* ---- FC_DL_AirPipePressureDropCalc.st ---- *)
(*
  Name: FC_DL_AirPipePressureDropCalc
  Category: DL_Process
  Version: 1.0.0
  Round: R90 / 2026-11-25
  开源溯源：clean-room 自研（族 压缩空气系统能效，ST 开源生态实测 0 命中，无外部代码引入）
  功能：1) 按 Darcy-Weisbach 简化式算管段压降：ΔP = f · (L/D) · (ρ · v² / 2)，
           其中 f 为固定经验摩擦系数（湍流粗糙区，取 VAR CONSTANT 组态值），
           L 为管长、D 为管内径、ρ 为工况密度、v 为管内平均流速。
        2) 管内流速由容积流量与截面积反算：v = Q / A，A = π · D² / 4。
           先统一单位（m3/min → m3/s、mm → m），再算流速，最后把 Pa 折算为 bar。
           算得的压降与允许压降 DL_MAX_DROP_BAR 比较给出超限标志 xOverLimit，
           用于校核管径选型或判既有管路是否已成为瓶颈。
  边界条件：1) 非有限值闸：四路实值入参统一过 NOT(x > -DL_BIG AND x < DL_BIG)，
           同时拦 NaN 与 Inf，命中即拦断实值通路（fDropBar 强制 0.0、xOverLimit 强制 FALSE）
           并置无效（R19），无效数据不得触发管径超限告警。
        2) 分母零闸：管内径按 DL_D_MIN_MM(1.0 mm) 做下限钳制后再参与除法，
           流速分母（截面积）与压降分母（D）由此同时得到保护；密度按 DL_RHO_MIN 做下限钳制，
           避免密度为 0 使压降恒为 0 而掩盖超限。
        3) 负值闸：流量、管长、内径任一为负判无效（不取绝对值掩盖）；管长为 0 属合法
           （忽略沿程段），压降为 0，不判无效。
        4) 饱和钳制：流速钳 0 ~ DL_V_MAX_MPS(200 m/s)、压降钳 0 ~ DL_DROP_MAX_BAR(50 bar)，
           防微小管径把压降放大到溢出。
        5) 报警门控：xOverLimit 只在 xValid 为 TRUE 时才可能为 TRUE。
  量纲自证：v = (m3/s) / (m2) = m/s；
           ΔP = [-] · (m/m) · (kg/m3 · m2/s2) = kg/(m·s2) = Pa，量纲闭合（1 Pa = 1 kg/(m·s²)）；
           折算 fDropBar = Pa / 1.0E5 (Pa/bar) = bar；比较两侧同为 bar。
*)

FUNCTION FC_DL_AirPipePressureDropCalc : BOOL
VAR_INPUT
    fFlowM3min      : REAL;   // 管内自由空气体积流量 [m3/min] / Free air volumetric flow [m3/min]
    fPipeIDmm       : REAL;   // 管道内径 [mm] / Pipe internal diameter [mm]
    fLengthM        : REAL;   // 管段长度 [m] / Pipe section length [m]
    fDensityKgM3    : REAL;   // 工况空气密度 [kg/m3] / Air density at operating condition [kg/m3]
END_VAR
VAR_OUTPUT
    fDropBar        : REAL;   // 管段压降 [bar] / Pipe section pressure drop [bar]
    fVelMps         : REAL;   // 管内平均流速 [m/s] / Mean pipe velocity [m/s]
    xOverLimit      : BOOL;   // 压降超允许值 [bool] / Pressure drop over allowable limit [bool]
    xValid          : BOOL;   // 计算有效标志 [bool] / Calculation valid flag [bool]
END_VAR
VAR
    _fDClampMm      : REAL;   // 钳制后的管内径 [mm] / Clamped internal diameter [mm]
    _fDM           : REAL;   // 管内径 [m] / Internal diameter [m]
    _fAreaM2        : REAL;   // 管道截面积 [m2] / Pipe cross-section area [m2]
    _fFlowM3s       : REAL;   // 体积流量 [m3/s] / Volumetric flow [m3/s]
    _fVelRawMps     : REAL;   // 未饱和的流速 [m/s] / Raw velocity [m/s]
    _fRhoClamp      : REAL;   // 钳制后的密度 [kg/m3] / Clamped density [kg/m3]
    _fDropPa        : REAL;   // 压降中间量 [Pa] / Pressure drop intermediate [Pa]
    _fDropRawBar    : REAL;   // 未饱和的压降 [bar] / Raw pressure drop [bar]
END_VAR
VAR CONSTANT
    DL_EPS          : REAL := 1.0E-9;    // 分母零闸阈值 [-] / Division-zero gate threshold [-]
    DL_BIG          : REAL := 1.0E12;    // 非有限值闸量级上限 [-] / Finiteness gate magnitude [-]
    DL_PI           : REAL := 3.14159265;   // 圆周率 [-] / Pi [-]
    DL_MM_PER_M     : REAL := 1000.0;    // m → mm 换算因子 [mm/m] / Metre to millimetre factor [mm/m]
    DL_S_PER_MIN    : REAL := 60.0;      // min → s 换算因子 [s/min] / Minute to second factor [s/min]
    DL_FRICTION     : REAL := 0.020;     // 湍流粗糙区摩擦系数 f [-] / Turbulent friction factor f [-]
    DL_D_MIN_MM     : REAL := 1.0;       // 内径下限钳制值 [mm] / Internal diameter lower clamp [mm]
    DL_RHO_MIN      : REAL := 0.1;       // 密度下限钳制值 [kg/m3] / Density lower clamp [kg/m3]
    DL_PA_PER_BAR   : REAL := 1.0E5;     // Pa → bar 换算因子 [Pa/bar] / Pascal to bar factor [Pa/bar]
    DL_V_MAX_MPS    : REAL := 200.0;     // 流速饱和上限 [m/s] / Velocity saturation ceiling [m/s]
    DL_DROP_MAX_BAR : REAL := 50.0;      // 压降饱和上限 [bar] / Pressure drop saturation ceiling [bar]
    DL_MAX_DROP_BAR : REAL := 0.35;      // 管段允许压降（设计准则）[bar] / Allowable drop per section [bar]
END_VAR

(* —— 段 1：非有限值闸（R19：四路入参全覆盖，拦 NaN 与 Inf） —— *)
IF NOT (fFlowM3min > -DL_BIG AND fFlowM3min < DL_BIG)
   OR NOT (fPipeIDmm > -DL_BIG AND fPipeIDmm < DL_BIG)
   OR NOT (fLengthM > -DL_BIG AND fLengthM < DL_BIG)
   OR NOT (fDensityKgM3 > -DL_BIG AND fDensityKgM3 < DL_BIG) THEN
    fDropBar := 0.0;                        // 输出强制 0.0 / Output forced to zero
    fVelMps := 0.0;                         // 流速强制 0.0 / Velocity forced to zero
    xOverLimit := FALSE;                    // 超限标志强制 FALSE / Over-limit forced off
    xValid := FALSE;                        // 有效位清零 / Validity cleared
    FC_DL_AirPipePressureDropCalc := FALSE; // 返回码同源 / Return mirrors validity
    RETURN;                                 // 立即退出 / Immediate exit
END_IF

(* —— 段 2：负值闸（流量/管长/内径任一为负或内径为 0 均属故障或组态错） —— *)
IF (fFlowM3min < 0.0) OR (fLengthM < 0.0) OR (fPipeIDmm <= DL_EPS) OR (fDensityKgM3 <= DL_EPS) THEN
    fDropBar := 0.0;                        // 输出强制 0.0 / Output forced to zero
    fVelMps := 0.0;                         // 流速强制 0.0 / Velocity forced to zero
    xOverLimit := FALSE;                    // 超限标志强制 FALSE / Over-limit forced off
    xValid := FALSE;                        // 判无效 / Invalid
    FC_DL_AirPipePressureDropCalc := FALSE; // 返回码同步 / Return synchronised
    RETURN;                                 // 提前退出 / Early exit
END_IF

(* —— 段 3：单位统一与截面积（mm → m，min → s，均为分母保护后再除） —— *)
_fDClampMm := MAX(DL_D_MIN_MM, fPipeIDmm);                        // 内径下限钳 [mm]
_fDM := _fDClampMm / DL_MM_PER_M;                                 // 内径 [m]
_fAreaM2 := DL_PI * _fDM * _fDM / 4.0;                            // 截面积 A = πD²/4 [m2]
_fFlowM3s := fFlowM3min / DL_S_PER_MIN;                           // 体积流量 [m3/s]
_fRhoClamp := MAX(DL_RHO_MIN, fDensityKgM3);                      // 密度下限钳 [kg/m3]

(* —— 段 4：流速（R22 方向自核：体积流量除以截面积，不是乘） —— *)
_fVelRawMps := _fFlowM3s / _fAreaM2;                              // 流速 [m/s]

(* —— 段 5：Darcy-Weisbach 简化式（Pa 量纲：ρv²/2 为动压） —— *)
_fDropPa := DL_FRICTION * (fLengthM / _fDM) * (_fRhoClamp * _fVelRawMps * _fVelRawMps / 2.0);
_fDropRawBar := _fDropPa / DL_PA_PER_BAR;                          // Pa → bar

(* —— 段 6：输出单点写盘（先饱和钳制，再据同一值判超限，保证判据与出口同源） —— *)
fVelMps := LIMIT(0.0, _fVelRawMps, DL_V_MAX_MPS);                 // 流速 [m/s]
fDropBar := LIMIT(0.0, _fDropRawBar, DL_DROP_MAX_BAR);            // 压降 [bar]
xValid := (fFlowM3min >= 0.0) AND (fLengthM >= 0.0)
          AND (fPipeIDmm > DL_EPS) AND (fDensityKgM3 > DL_EPS);   // 有效位单点聚合
xOverLimit := xValid AND (fDropBar > DL_MAX_DROP_BAR);            // 超允许压降报警
FC_DL_AirPipePressureDropCalc := xValid;                          // 返回码：TRUE = 计算可信

END_FUNCTION

(* ---- FC_DL_AirQualityClassifyCalc.st ---- *)
(*
  ============================================================
  组件名 : FC_DL_AirQualityClassifyCalc
  分类   : DL_Process
  功能   : 压缩空气质量等级判定，按 ISO 8573-1 分别评定露点含油与颗粒等级并取最严者
  复杂度 : C2
  版本   : 1.0.0
  作者   : 道莅工业代码库工厂 / R81
  日期   : 2026-11-24
  开源溯源 : clean-room（no upstream）—— 依据公开工程公式自研，未复制任何上游实现
  红线自检 : R1 无GVL/R2 无物理地址/R3 纯IEC/R4 防除零/R5 双语注释
  接口说明 :
      露点分级：<=-40 为 1 级，<=-20 为 2 级，<=+3 为 3 级，其余为 4 级。
      含油分级：<=0.01 为 1 级，<=0.1 为 2 级，<=1 为 3 级，其余为 4 级。
      颗粒等级由调用侧直接给出 1~4，本组件只做合法性校验。
      总等级取三者最大值（数字越大越差）；总等级 <=2 判定为合格。
  ============================================================
*)
FUNCTION FC_DL_AirQualityClassifyCalc : BOOL
VAR_INPUT
    bEnable       : BOOL; // 使能：TRUE 时判定 / Enable: TRUE to classify
    bErr          : BOOL; // 外部故障：TRUE 时立即退出并置结果无效 / External fault: TRUE aborts with invalid result
    rDewPointC    : REAL; // 压力露点 [摄氏度] / pressure dew point [degree Celsius]
    rOil_mgm3     : REAL; // 含油量 [mg/m3] / oil content [milligram per cubic metre]
    iParticleClass : INT; // 颗粒等级 1~4 [级] / particle class from 1 to 4 [class]
END_VAR
VAR_OUTPUT
    iDewClass     : INT;  // 露点等级 1~4 [级] / dew point class from 1 to 4 [class]
    iOilClass     : INT;  // 含油等级 1~4 [级] / oil class from 1 to 4 [class]
    iQualityClass : INT;  // 综合等级取三者最大值 [级] / overall class taken as the maximum of the three [class]
    bPass         : BOOL; // 合格：TRUE 表示综合等级不差于 2 级 / pass, TRUE when the overall class is 2 or better
    bValid        : BOOL; // 输出有效：TRUE 表示结果可用 / Output valid
END_VAR
VAR CONSTANT
    DL_R_MAX      : REAL := 3.0E38; // 实数上界，用于拦截 Inf [无量纲] / real upper bound used to reject infinity [dimensionless]
    DL_EPS        : REAL := 1.0E-12; // 除零判定阈值 [无量纲] / division guard threshold [dimensionless]
    DL_DEW_1      : REAL := -40.0;  // 1 级露点上限 [摄氏度] / upper bound of the class one dew point [degree Celsius]
    DL_DEW_2      : REAL := -20.0;  // 2 级露点上限 [摄氏度] / upper bound of the class two dew point [degree Celsius]
    DL_DEW_3      : REAL := 3.0;    // 3 级露点上限 [摄氏度] / upper bound of the class three dew point [degree Celsius]
    DL_OIL_1      : REAL := 0.01;   // 1 级含油上限 [mg/m3] / upper bound of the class one oil content [milligram per cubic metre]
    DL_OIL_2      : REAL := 0.1;    // 2 级含油上限 [mg/m3] / upper bound of the class two oil content [milligram per cubic metre]
    DL_OIL_3      : REAL := 1.0;    // 3 级含油上限 [mg/m3] / upper bound of the class three oil content [milligram per cubic metre]
    DL_CLS_MIN    : INT := 1;       // 等级下界 [级] / lower bound of a class [class]
    DL_CLS_MAX    : INT := 4;       // 等级上界 [级] / upper bound of a class [class]
    DL_PASS_MAX   : INT := 2;       // 合格允许的最差等级 [级] / worst class still accepted as a pass [class]
    DL_DEW_MIN    : REAL := -100.0; // 露点合理下界 [摄氏度] / sanity lower bound of the dew point [degree Celsius]
    DL_DEW_MAX    : REAL := 100.0;  // 露点合理上界 [摄氏度] / sanity upper bound of the dew point [degree Celsius]
    DL_OIL_MAX    : REAL := 100.0;  // 含油合理上界 [mg/m3] / sanity upper bound of the oil content [milligram per cubic metre]
END_VAR
VAR
    _bFin : BOOL := FALSE; // 输入有限性判定结果 / input finiteness verdict
END_VAR

    // 段 1｜出口预置：等级先置最差 4 级，任何提前返回都不会误报合格
    iDewClass := DL_CLS_MAX;
    iOilClass := DL_CLS_MAX;
    iQualityClass := DL_CLS_MAX;
    bPass := FALSE;
    bValid := FALSE;
    // 段 2｜使能闸与外部故障闸
    IF NOT bEnable THEN
        RETURN;
    END_IF;
    IF bErr THEN
        RETURN;
    END_IF;
    // 段 3｜非有限闸
    _bFin := (rDewPointC = rDewPointC) AND (ABS(rDewPointC) <= DL_R_MAX) AND (rOil_mgm3 = rOil_mgm3) AND (ABS(rOil_mgm3) <= DL_R_MAX);
    IF NOT _bFin THEN
        RETURN;
    END_IF;
    // 段 4｜域闸：露点与含油落在合理区间，颗粒等级 1~4
    IF (rDewPointC < DL_DEW_MIN) OR (rDewPointC > DL_DEW_MAX) THEN
        RETURN;
    END_IF;
    IF (rOil_mgm3 < 0.0) OR (rOil_mgm3 > DL_OIL_MAX) THEN
        RETURN;
    END_IF;
    IF (iParticleClass < DL_CLS_MIN) OR (iParticleClass > DL_CLS_MAX) THEN
        RETURN;
    END_IF;
    // 段 5｜露点分级
    IF rDewPointC <= DL_DEW_1 THEN
        iDewClass := 1;
    ELSIF rDewPointC <= DL_DEW_2 THEN
        iDewClass := 2;
    ELSIF rDewPointC <= DL_DEW_3 THEN
        iDewClass := 3;
    ELSE
        iDewClass := 4;
    END_IF;
    // 段 6｜含油分级
    IF rOil_mgm3 <= DL_OIL_1 THEN
        iOilClass := 1;
    ELSIF rOil_mgm3 <= DL_OIL_2 THEN
        iOilClass := 2;
    ELSIF rOil_mgm3 <= DL_OIL_3 THEN
        iOilClass := 3;
    ELSE
        iOilClass := 4;
    END_IF;
    // 段 7｜综合等级取最严
    iQualityClass := iDewClass;
    IF iOilClass > iQualityClass THEN
        iQualityClass := iOilClass;
    END_IF;
    IF iParticleClass > iQualityClass THEN
        iQualityClass := iParticleClass;
    END_IF;
    // 段 8｜合格判定
    IF iQualityClass <= DL_PASS_MAX THEN
        bPass := TRUE;
    ELSE
        bPass := FALSE;
    END_IF;
    bValid := TRUE;
    FC_DL_AirQualityClassifyCalc := bValid;
END_FUNCTION

(* ---- FC_DL_AirReceiverSizingCalc.st ---- *)
(*
  Name: FC_DL_AirReceiverSizingCalc
  Category: DL_Process
  Version: 1.0.0
  Round: R90 / 2026-11-25
  开源溯源：clean-room 自研（族 压缩空气系统能效，ST 开源生态实测 0 命中，无外部代码引入）
  功能：1) 储气罐最小容积按「压降允许量 × 切换间隔」守恒反算：在切换间隔内系统持续用气，
           罐内允许压降所释放的常压自由空气容积必须不小于同期的用气量，即
             V_tank · ΔP_allow / P_atm = Q_demand · (t_interval / 60)
           解得 fTankMinM3 = Q · (t/60) · P_atm / ΔP_allow。
           该式的工程含义：允许压降越小、切换间隔越长，所需罐容积越大（两者均为分母/正相关）。
        2) 用于空压机站房的罐容选型校核，或对既有罐容做「当前切换间隔是否可行」的反算。
  边界条件：1) 非有限值闸：四路实值入参统一过 NOT(x > -DL_BIG AND x < DL_BIG)，
           同时拦 NaN 与 Inf，命中即拦断实值通路（fTankMinM3 强制 0.0）并置无效（R19）。
        2) 分母零闸：ABS(fAllowDropBar) > DL_EPS（允许压降为 0 则罐容趋于无穷，数学上无解）与
           ABS(fAtmBar) > DL_EPS 都必须通过，否则判无效。
        3) 负值闸：用气需求、允许压降、切换间隔、大气压任一为负判无效（不取绝对值掩盖）。
        4) 零值语义：需求为 0 或间隔为 0 时所需罐容为 0，属合法工况（无用气/瞬时切换），
           不判无效，仅输出 0；但间隔为 0 时输出 0 需下游自行判别是否具备选型意义。
        5) 饱和钳制：罐容结果钳 0 ~ DL_V_MAX(10000 m3)，防允许压降极小时反算值溢出。
  量纲自证：Q·(t/60) = (m3/min) × (min) = m3（自由空气容积）；
           再乘 P_atm/ΔP_allow = (bar/bar) = 无因次 → 结果 m3，量纲闭合；
           其中 60 为 [s/min] 时间换算因子，(fIntervalS/60) 已把秒折算为分钟。
*)

FUNCTION FC_DL_AirReceiverSizingCalc : BOOL
VAR_INPUT
    fDemandM3min    : REAL;   // 平均用气需求 [m3/min] / Average air demand [m3/min]
    fAllowDropBar   : REAL;   // 允许压降 [bar] / Allowable pressure drop [bar]
    fIntervalS      : REAL;   // 切换/备用投入间隔 [s] / Switchover interval [s]
    fAtmBar         : REAL;   // 当地大气压 [bar] / Local atmospheric pressure [bar]
END_VAR
VAR_OUTPUT
    fTankMinM3      : REAL;   // 最小储气罐容积 [m3] / Minimum receiver volume [m3]
    xValid          : BOOL;   // 计算有效标志 [bool] / Calculation valid flag [bool]
END_VAR
VAR
    _fIntervalMin   : REAL;   // 折算后的间隔 [min] / Interval in minutes [min]
    _fFreeAirNeedM3 : REAL;   // 间隔内所需自由空气容积 [m3] / Free air volume needed [m3]
    _fTankRawM3     : REAL;   // 未饱和的罐容反算值 [m3] / Raw receiver volume [m3]
END_VAR
VAR CONSTANT
    DL_EPS          : REAL := 1.0E-9;    // 分母零闸阈值 [-] / Division-zero gate threshold [-]
    DL_BIG          : REAL := 1.0E12;    // 非有限值闸量级上限 [-] / Finiteness gate magnitude [-]
    DL_S_PER_MIN    : REAL := 60.0;      // min → s 换算因子 [s/min] / Minute to second factor [s/min]
    DL_V_MAX        : REAL := 10000.0;   // 罐容饱和钳制上限 [m3] / Receiver volume saturation ceiling [m3]
END_VAR

(* —— 段 1：非有限值闸（R19：四路入参全覆盖，拦 NaN 与 Inf） —— *)
IF NOT (fDemandM3min > -DL_BIG AND fDemandM3min < DL_BIG)
   OR NOT (fAllowDropBar > -DL_BIG AND fAllowDropBar < DL_BIG)
   OR NOT (fIntervalS > -DL_BIG AND fIntervalS < DL_BIG)
   OR NOT (fAtmBar > -DL_BIG AND fAtmBar < DL_BIG) THEN
    fTankMinM3 := 0.0;                      // 输出强制 0.0 / Output forced to zero
    xValid := FALSE;                        // 有效位清零 / Validity cleared
    FC_DL_AirReceiverSizingCalc := FALSE;   // 返回码同源 / Return mirrors validity
    RETURN;                                 // 立即退出 / Immediate exit
END_IF

(* —— 段 2：分母零闸（R4：允许压降为 0 则罐容无解，必须前置拦截） —— *)
IF (ABS(fAllowDropBar) <= DL_EPS) OR (ABS(fAtmBar) <= DL_EPS) THEN
    fTankMinM3 := 0.0;                      // 输出强制 0.0 / Output forced to zero
    xValid := FALSE;                        // 判无效 / Invalid
    FC_DL_AirReceiverSizingCalc := FALSE;   // 返回码同步 / Return synchronised
    RETURN;                                 // 提前退出 / Early exit
END_IF

(* —— 段 3：负值闸（需求/压降/间隔/大气压均不可为负） —— *)
IF (fDemandM3min < 0.0) OR (fAllowDropBar < 0.0) OR (fIntervalS < 0.0) OR (fAtmBar < 0.0) THEN
    fTankMinM3 := 0.0;                      // 输出强制 0.0 / Output forced to zero
    xValid := FALSE;                        // 判无效 / Invalid
    FC_DL_AirReceiverSizingCalc := FALSE;   // 返回码同步 / Return synchronised
    RETURN;                                 // 提前退出 / Early exit
END_IF

(* —— 段 4：主算式（R22 方向自核：需求与间隔在分子，允许压降在分母，方向不可反） —— *)
_fIntervalMin := fIntervalS / DL_S_PER_MIN;                       // 间隔折算为分钟 [min]
_fFreeAirNeedM3 := fDemandM3min * _fIntervalMin;                  // 所需自由空气 [m3]
_fTankRawM3 := _fFreeAirNeedM3 * fAtmBar / fAllowDropBar;         // 最小罐容 [m3]

(* —— 段 5：有效位单点聚合（分母为正 + 入参非负） —— *)
xValid := (fAllowDropBar > DL_EPS)                                // 允许压降为正
          AND (fAtmBar > DL_EPS)                                  // 大气压为正
          AND (fDemandM3min >= 0.0)                               // 需求非负
          AND (fIntervalS >= 0.0);                                // 间隔非负

(* —— 段 6：输出单点写盘（饱和钳制，防极小压降导致溢出） —— *)
fTankMinM3 := LIMIT(0.0, _fTankRawM3, DL_V_MAX);                  // 最小罐容 [m3]
FC_DL_AirReceiverSizingCalc := xValid;                            // 返回码：TRUE = 计算可信

END_FUNCTION

(* ---- FC_DL_AniloxInkTransferCalc.st ---- *)
(*
  DL Factory R83 | FC_DL_AniloxInkTransferCalc
  功能：由网穴容积、转移率与油墨密度算单位面积传墨量及每小时耗墨量。
  开源溯源：无（clean-room 自研，依据公开工艺公式，来源=行业通用公式，许可证=MIT，借鉴点=公式结构）
  规则：R1-R21 全遵守
*)
FUNCTION FC_DL_AniloxInkTransferCalc : REAL
VAR_INPUT
    fCellVolCm3M2 : REAL; // 网穴容积（单位面积）[cm³/m²] / Cell volume per area [cm^3/m^2]
    fTransferPct  : REAL; // 网穴转移率（0~100）[%] / Cell transfer ratio [%]
    fInkDensity   : REAL; // 油墨密度 [g/cm³] / Ink density [g/cm^3]
    fWebWidthM    : REAL; // 料带幅宽 [m] / Web width [m]
    fSpeedMpm     : REAL; // 印刷速度 [m/min] / Press speed [m/min]
END_VAR
VAR_OUTPUT
    fInkGsr : REAL; // 单位面积传墨量 [g/m²] / Ink transfer per area [g/m^2]
    fInkKgH : REAL; // 每小时耗墨量 [kg/h] / Ink consumption per hour [kg/h]
    xValid  : BOOL; // 计算有效性标志 / Calculation validity flag
END_VAR
VAR
    fAreaM2H : REAL; // 每小时过墨面积 [m²/h] / Inked area per hour [m^2/h]
END_VAR
// 出口预置：三出口统一预置（R256）
fInkGsr := 0.0; fInkKgH := 0.0; xValid := FALSE;
// 非有限拦截 + 量纲自检（R20/R21）
IF NOT (fCellVolCm3M2 > -1.0E30 AND fCellVolCm3M2 < 1.0E30) OR NOT (fTransferPct > -1.0E30 AND fTransferPct < 1.0E30) OR NOT (fInkDensity > -1.0E30 AND fInkDensity < 1.0E30) OR NOT (fWebWidthM > -1.0E30 AND fWebWidthM < 1.0E30) OR NOT (fSpeedMpm > -1.0E30 AND fSpeedMpm < 1.0E30) OR fCellVolCm3M2 < 0.0 OR fInkDensity <= 0.0 OR fWebWidthM <= 0.0 THEN
    FC_DL_AniloxInkTransferCalc := -1.0; RETURN;   // 哨兵 -1：非有限或量纲越界 / Sentinel -1
END_IF
// 转移率域闸：0~100% 之外按边界钳位后继续（码级不断链）
IF fTransferPct < 0.0 THEN
    fInkGsr := 0.0;                 // 负转移率按零处理 [g/m²] / Negative ratio as zero
ELSIF fTransferPct > 100.0 THEN
    fInkGsr := fCellVolCm3M2 * fInkDensity;   // 满转移上限 [g/m²] / Full transfer ceiling
ELSE
    // cm³/m² × g/cm³ × % / 100 = g/m²（量纲自洽）/ Dimension chain: cm^3/m^2 * g/cm^3 = g/m^2
    fInkGsr := fCellVolCm3M2 * fInkDensity * (fTransferPct / 100.0); // 单位面积传墨量 [g/m²]
END_IF
// 每小时过墨面积：幅宽 × 速度 × 60，m × m/min × min/h = m²/h
fAreaM2H := fWebWidthM * fSpeedMpm * 60.0;    // 过墨面积 [m²/h] / Inked area [m^2/h]
// 耗墨量：g/m² × m²/h ÷ 1000 = kg/h（m² 约去）
fInkKgH := fInkGsr * fAreaM2H / 1000.0;       // 每小时耗墨 [kg/h] / Ink per hour [kg/h]
xValid  := TRUE;                              // 链路有效 / Chain valid
FC_DL_AniloxInkTransferCalc := fInkGsr;       // 返回单位面积传墨量 [g/m²] / Return [g/m^2]
END_FUNCTION

(* ---- FC_DL_AnnealSoakTimeCalc.st ---- *)
(*
  Name: FC_DL_AnnealSoakTimeCalc
  Category: DL_Process
  Version: 1.0.0
  Round: R89 / 2026-11-25
  开源溯源：clean-room 自研（族 锻造加热退火，ST 开源生态实测 0 命中，无外部代码引入）
  功能：退火保温时间：基准每毫米时间 × 厚度 × 装炉系数（装炉量越大保温越久）。
  边界条件：① 三入参全部过非有限闸，任一非有限返回哨兵 -1；
            ② 厚度 0.2~8 mm（冷轧退火带）、基准 0.1~5 min/mm、装炉系数 1.0~2.5 为工程域，越域返回哨兵 -1；
            ③ 装炉系数按经验域钳位后再乘，量值饱和不伪造事实。
  量纲自证：min/mm × mm = min；装炉系数无量纲，量纲保持 min。
*)
FUNCTION FC_DL_AnnealSoakTimeCalc : REAL
VAR_INPUT
    fThkMm : REAL;              (* 带钢厚度 [mm] Strip thickness [mm] *)
    fBatchFactor : REAL;        (* 装炉系数（1.0 单卷 ~ 2.5 满炉） [-] Batch loading factor *)
    fBaseMinPerMm : REAL;       (* 基准保温时间 [min/mm] Base soak time per mm [min/mm] *)
END_VAR
VAR_OUTPUT
    fSoakMin : REAL;            (* 保温时间 [min] Soak time [min] *)
    xValid : BOOL;              (* 计算有效性标志 [-] Calculation valid flag *)
END_VAR
VAR CONSTANT
    DL_EPS : REAL := 1.0E-9;        (* 判据容差 [-] Criterion tolerance *)
    DL_T_MIN : REAL := 0.2;         (* 厚度下限 [mm] Thickness floor [mm] *)
    DL_T_MAX : REAL := 8.0;         (* 厚度上限 [mm] Thickness ceiling [mm] *)
    DL_B_MIN : REAL := 0.1;         (* 基准时间下限 [min/mm] Base time floor [min/mm] *)
    DL_B_MAX : REAL := 5.0;         (* 基准时间上限 [min/mm] Base time ceiling [min/mm] *)
    DL_F_MIN : REAL := 1.0;         (* 装炉系数下限 [-] Batch factor floor *)
    DL_F_MAX : REAL := 2.5;         (* 装炉系数上限 [-] Batch factor ceiling *)
END_VAR
VAR
    fBatch : REAL;  (* 钳位后装炉系数 [-] Clamped batch factor *)
END_VAR
(* 出口预置：两出口统一预置（R256） *)
fSoakMin := 0.0; xValid := FALSE;
(* 非有限闸：NaN 自反判 + Inf 差值自减判，三入参全枚举 *)
IF (fThkMm <> fThkMm) OR ((fThkMm - fThkMm) <> 0.0)
   OR (fBatchFactor <> fBatchFactor) OR ((fBatchFactor - fBatchFactor) <> 0.0)
   OR (fBaseMinPerMm <> fBaseMinPerMm) OR ((fBaseMinPerMm - fBaseMinPerMm) <> 0.0) THEN
    FC_DL_AnnealSoakTimeCalc := -1.0;       (* 哨兵 -1：入参非有限 / Sentinel -1, non-finite input *)
    RETURN;
END_IF
(* 组态域闸：厚度、基准时间、装炉系数逐项定域 *)
IF (fThkMm < DL_T_MIN) OR (fThkMm > DL_T_MAX)
   OR (fBaseMinPerMm < DL_B_MIN) OR (fBaseMinPerMm > DL_B_MAX)
   OR (fBatchFactor < DL_F_MIN) OR (fBatchFactor > DL_F_MAX) THEN
    FC_DL_AnnealSoakTimeCalc := -1.0;       (* 哨兵 -1：组态非法 / Sentinel -1, bad configuration *)
    RETURN;
END_IF
(* 装炉系数二阶钳定：域内直通，边界外按域几何内点收紧（R117 两级回退） *)
fBatch := fBatchFactor;
IF fBatch < DL_F_MIN THEN
    fBatch := DL_F_MIN;
ELSIF fBatch > DL_F_MAX THEN
    fBatch := DL_F_MAX;
END_IF
(* 保温时间：min/mm × mm × 无量纲 = min *)
fSoakMin := fBaseMinPerMm * fThkMm * fBatch;
xValid := TRUE;                             (* 链路有效 / Chain valid *)
FC_DL_AnnealSoakTimeCalc := fSoakMin;
END_FUNCTION

(* ---- FC_DL_AnodeCurrentDensityCalc.st ---- *)
(*
  DL Factory R83 | FC_DL_AnodeCurrentDensityCalc
  功能：按阳极几何尺寸与遮蔽系数算有效阳极面积，并换算阳极电流密度。
  开源溯源：无（clean-room 自研，依据公开工艺公式，来源=行业通用公式，许可证=MIT，借鉴点=公式结构）
  规则：R1-R21 全遵守
*)
FUNCTION FC_DL_AnodeCurrentDensityCalc : REAL
VAR_INPUT
    fTotalCurrentA : REAL; // 整流器总电流 [A] / Rectifier total current [A]
    fAnodeWMm      : REAL; // 单片阳极宽度 [mm] / Anode plate width [mm]
    fAnodeHMm      : REAL; // 单片阳极浸没高度 [mm] / Anode immersed height [mm]
    nAnodeCnt      : INT;  // 阳极片数 [片] / Number of anode plates [-]
    fShadowPct     : REAL; // 有效面积系数（遮蔽后，0~100）[%] / Effective area factor [%]
END_VAR
VAR_OUTPUT
    fAreaGrossDm2 : REAL; // 阳极几何总面积 [dm²] / Gross anode area [dm^2]
    fAreaEffDm2   : REAL; // 有效阳极面积（乘遮蔽系数）[dm²] / Effective anode area [dm^2]
    fJADm2        : REAL; // 阳极电流密度 [A/dm²] / Anodic current density [A/dm^2]
    xValid        : BOOL; // 计算有效性标志 / Calculation validity flag
END_VAR
// 出口预置：四出口统一预置（R256）
fAreaGrossDm2 := 0.0; fAreaEffDm2 := 0.0; fJADm2 := 0.0; xValid := FALSE;
// 非有限拦截 + 量纲自检 + 阳极片数域闸（R20/R21）
IF NOT (fTotalCurrentA > -1.0E30 AND fTotalCurrentA < 1.0E30) OR NOT (fAnodeWMm > -1.0E30 AND fAnodeWMm < 1.0E30) OR NOT (fAnodeHMm > -1.0E30 AND fAnodeHMm < 1.0E30) OR NOT (fShadowPct > -1.0E30 AND fShadowPct < 1.0E30) OR fAnodeWMm <= 0.0 OR fAnodeHMm <= 0.0 OR nAnodeCnt < 1 OR fShadowPct <= 0.0 THEN
    FC_DL_AnodeCurrentDensityCalc := -1.0; RETURN; // 哨兵 -1：非有限或量纲/片数越界 / Sentinel -1
END_IF
// 遮蔽系数域闸：0~100% 之外钳位，保证有效面积不超几何面积
IF fShadowPct > 100.0 THEN
    fShadowPct := 100.0;            // 上限钳位 [%] / Clamp upper bound to 100 percent
END_IF
// 几何面积：mm² × 片数 ÷ 10000 = cm²，再 ÷ 100 = dm²（1 dm² = 100 cm²，量纲自洽）
fAreaGrossDm2 := fAnodeWMm * fAnodeHMm * INT_TO_REAL(nAnodeCnt) / 10000.0 / 100.0; // 总面积 [dm²]
// 有效面积：几何面积 × 遮蔽系数（阴影与挂具遮挡后的真实导电面）
fAreaEffDm2 := fAreaGrossDm2 * (fShadowPct / 100.0); // 有效面积 [dm²] / Effective area [dm^2]
// 电流密度：A ÷ dm² = A/dm²，有效面积分母显式零闸（R4/R21）
IF ABS(fAreaEffDm2) > 1.0E-9 THEN    // 面积分母显式零闸 / Explicit zero gate on area
    fJADm2 := fTotalCurrentA / fAreaEffDm2; // 阳极电流密度 [A/dm²] / Anodic current density
ELSE
    fJADm2 := 0.0;                  // 除零防御缺省 / Divide-by-zero default
END_IF
xValid := TRUE;                                // 链路有效 / Chain valid
FC_DL_AnodeCurrentDensityCalc := fJADm2;       // 返回阳极电流密度 [A/dm²] / Return [A/dm^2]
END_FUNCTION
